(* IEC 61131-3 sources: Industry-PLC-LLM/data/PLCBEAD_repo/PLCBEAD_PLCEmbed-main/PLC-BEAD/Source/OpenPLCv3 (part 4) *)

(* ---- CYCLE_TIME.ST ---- *)
FUNCTION_BLOCK T_PLC_MS_block
	VAR_OUTPUT
		T_PLC_MS :	UDINT;
	END_VAR

	VAR_EXTERNAL
		PLC_TICKS_PER_SEC :	INT;
		PLC_SYS_TICK_CNT :	DINT;
	END_VAR

	VAR
		debug :	BOOL;(*Debug-Mode ON / OFF*)
		N :	INT;(*Debug-Faktor*)
		Offset :	UDINT;(*Debug-Offset*)
		temp :	DWORD := DWORD#1;(*Debug-Offset*)
		mode :	BOOL;(*modus*)
		faktor :	UDINT;(*Systemtakt-Faktor*)
		init :	BOOL;
		v_plc_ticks_per_sec :	UDINT;
		base :	UDINT := UDINT#1000;
	END_VAR

	IF init = FALSE THEN
		v_plc_ticks_per_sec := INT_TO_UDINT(PLC_TICKS_PER_SEC);
		IF v_plc_ticks_per_sec = UDINT#1024 THEN
			faktor := UDINT#1;
			mode := FALSE;
		ELSIF v_plc_ticks_per_sec > UDINT#0 THEN
			IF v_plc_ticks_per_sec <= base THEN
				faktor := base / v_plc_ticks_per_sec;
				mode := FALSE;
			ELSE
				faktor := v_plc_ticks_per_sec / base;
				mode := TRUE;
			END_IF;
		ELSE
			faktor := UDINT#1;
		END_IF;
		init := TRUE;
	END_IF;

	IF mode THEN
		T_PLC_MS := DINT_TO_UDINT(PLC_SYS_TICK_CNT) / faktor;
	ELSE
		T_PLC_MS := DINT_TO_UDINT(PLC_SYS_TICK_CNT) * faktor;
	END_IF;

	IF debug THEN
		T_PLC_MS := (DWORD_TO_UDINT(SHL(UDINT_TO_DWORD(T_PLC_MS),N) OR SHL(temp,N)) - UDINT#1) + Offset;
	END_IF;

END_FUNCTION_BLOCK

FUNCTION_BLOCK CYCLE_TIME
	VAR_INPUT
		RST :	BOOL;
	END_VAR

	VAR_OUTPUT
		CT_MIN :	TIME := t#0s;
		CT_MAX :	TIME := t#0s;
		CT_LAST :	TIME;
		SYSTIME :	TIME;
		SYSDAYS :	INT;
		CYCLES :	DWORD;
	END_VAR

	VAR
		last_cycle :	TIME;
		tx :	TIME;
		init :	BOOL;
		T_PLC_MS :	T_PLC_MS_block;
	END_VAR

	T_PLC_MS();
	tx:= UDINT_TO_TIME(T_PLC_MS.T_PLC_MS) - last_cycle;

	IF rst THEN
		ct_min := t#10h;
		ct_max := t#0ms;
		cycles := DWORD#0;
	ELSIF last_cycle > t#0s THEN
		IF tx < ct_min THEN ct_min := tx;
		ELSIF tx > ct_max THEN ct_max := tx;
		END_IF;
		ct_last := tx;
	ELSIF ct_min = t#0s THEN
		ct_min := t#0s - t#1ms;
	END_IF;
	IF init THEN
		systime := systime + tx;
			IF systime >= t#1d THEN
				systime := systime - t#1d;
				sysdays := sysdays + 1;
			END_IF;
	END_IF;
	init := TRUE;
	last_cycle := last_cycle + tx;
	cycles := UDINT_TO_DWORD(DWORD_TO_UDINT(cycles) + UDINT#1);

END_FUNCTION_BLOCK

PROGRAM program0
  VAR
	RST :	BOOL;

	CT_MIN  :	TIME;
	CT_MAX  :	TIME;
	CT_LAST :	TIME;
	SYSTIME :	TIME;
	SYSDAYS :	INT;
	CYCLES  :	DWORD;

	func_block : CYCLE_TIME;
  END_VAR
	func_block.RST   :=RST ;
	func_block();
	CT_MIN := func_block.CT_MIN ;
	CT_MAX := func_block.CT_MAX ;
	CT_LAST:= func_block.CT_LAST;
	SYSTIME:= func_block.SYSTIME;
	SYSDAYS:= func_block.SYSDAYS;
	CYCLES := func_block.CYCLES ;
END_PROGRAM

CONFIGURATION Config0
	VAR_GLOBAL
		PLC_TICKS_PER_SEC :	INT;
		PLC_SYS_TICK_CNT :	DINT;
	END_VAR

  	RESOURCE Res0 ON PLC
    	TASK task0(INTERVAL := T#20ms,PRIORITY := 0);
    	PROGRAM instance0 WITH task0 : program0;
  	END_RESOURCE
END_CONFIGURATION

(* ---- D_TRIG.ST ---- *)
FUNCTION_BLOCK D_TRIG
	VAR_INPUT
		IN :	DWORD;
	END_VAR

	VAR_OUTPUT
		Q :	BOOL;
		X :	DWORD;
	END_VAR

	VAR
		last_in :	DWORD;
	END_VAR

	Q := in <> last_in;
	X := UDINT_TO_DWORD(DWORD_TO_UDINT(in) - DWORD_TO_UDINT(last_in));
	last_in := in;
END_FUNCTION_BLOCK

PROGRAM program0
  VAR
	IN :	DWORD;

	Q :	BOOL;
	X :	DWORD;

	func_block : D_TRIG;
  END_VAR
	func_block.IN  := IN;
	func_block();
	Q := func_block.Q;
	X := func_block.X;
END_PROGRAM

CONFIGURATION Config0
  RESOURCE Res0 ON PLC
    TASK task0(INTERVAL := T#20ms,PRIORITY := 0);
    PROGRAM instance0 WITH task0 : program0;
  END_RESOURCE
END_CONFIGURATION

(* ---- DATE_TO_STRING.ST ---- *)
FUNCTION YEAR_OF_DATE:INT
	VAR_INPUT
		IDATE :	UDINT;
	END_VAR

	YEAR_OF_DATE := UDINT_TO_INT((idate+UDINT#43200) / UDINT#31557600 + UDINT#1970);
END_FUNCTION

FUNCTION DAY_OF_YEAR:INT
	VAR_INPUT
		IDATE :	UDINT;
	END_VAR

	DAY_OF_YEAR := UDINT_TO_INT(((idate) / UDINT#86400) MOD UDINT#1461);
	IF DAY_OF_YEAR > 729 THEN
		IF DAY_OF_YEAR > 1095 THEN DAY_OF_YEAR := DAY_OF_YEAR - 1095; ELSE DAY_OF_YEAR := DAY_OF_YEAR - 729; END_IF;
	ELSIF DAY_OF_YEAR > 364 THEN
		DAY_OF_YEAR := DAY_OF_YEAR - 364;
	ELSE
		DAY_OF_YEAR := DAY_OF_YEAR + 1;
	END_IF;
END_FUNCTION

FUNCTION LEAP_OF_DATE:BOOL

	VAR_INPUT
		IDATE :	UDINT;
	END_VAR

	LEAP_OF_DATE := SHL(UDINT_TO_DWORD((idate + UDINT#43200) / UDINT#31557600), 30) = DWORD#16#80000000;
END_FUNCTION

FUNCTION MONTH_OF_DATE:INT

	VAR_INPUT
		IDATE :	UDINT;
	END_VAR

	MONTH_OF_DATE := DAY_OF_YEAR(idate);
	IF MONTH_OF_DATE < 32 THEN
		MONTH_OF_DATE := 1;
	ELSIF LEAP_OF_DATE((IDATE)) THEN
		MONTH_OF_DATE := (MONTH_OF_DATE * 53 + 1668) / 1623;
	ELSE
		MONTH_OF_DATE := (MONTH_OF_DATE * 53 + 1700) / 1620;
	END_IF;
END_FUNCTION

FUNCTION DAY_OF_MONTH:INT
	VAR_INPUT
		IDATE :	UDINT;
	END_VAR

	day_of_month := day_of_year(idate);

	IF leap_of_Date((idate)) THEN
		CASE day_of_month OF
			32..60	:	day_of_month := day_of_month - 31;
			61..91	:	day_of_month := day_of_month - 60;
			92..121 :	day_of_month := day_of_month - 91;
			122..152:	day_of_month := day_of_month - 121;
			153..182:	day_of_month := day_of_month - 152;
			183..213:	day_of_month := day_of_month - 182;
			214..244:	day_of_month := day_of_month - 213;
			245..274:	day_of_month := day_of_month - 244;
			275..305:	day_of_month := day_of_month - 274;
			306..335:	day_of_month := day_of_month - 305;
			336..366:	day_of_month := day_of_month - 335;
		END_CASE;
	ELSE
		CASE day_of_month OF
			32..59	:	day_of_month := day_of_month - 31;
			60..90	:	day_of_month := day_of_month - 59;
			91..120 :	day_of_month := day_of_month - 90;
			121..151:	day_of_month := day_of_month - 120;
			152..181:	day_of_month := day_of_month - 151;
			182..212:	day_of_month := day_of_month - 181;
			213..243:	day_of_month := day_of_month - 212;
			244..273:	day_of_month := day_of_month - 243;
			274..304:	day_of_month := day_of_month - 273;
			305..334:	day_of_month := day_of_month - 304;
			335..365:	day_of_month := day_of_month - 334;
		END_CASE;
	END_IF;
END_FUNCTION

FUNCTION_BLOCK DATE_TO_STRING2
	VAR_INPUT
		IDATE :	UDINT;
	END_VAR

	VAR_OUTPUT
		DATE_STRING :	STRING;
	END_VAR

	VAR
		st_tmp1 :	STRING;
	END_VAR

	st_tmp1 := CONCAT(INT_TO_STRING(YEAR_OF_DATE(IDATE)),INT_TO_STRING(MONTH_OF_DATE(IDATE)));
	DATE_STRING := CONCAT(st_tmp1,INT_TO_STRING(day_of_month(IDATE)));
END_FUNCTION_BLOCK

PROGRAM program0
  VAR
    LocalVar0 : UDINT;
	LocalOUT  : STRING;
	func_block : DATE_TO_STRING2;
  END_VAR
	func_block.IDATE  := LocalVar0;
	func_block();
	LocalOUT := func_block.DATE_STRING;
END_PROGRAM

CONFIGURATION Config0
  RESOURCE Res0 ON PLC
    TASK task0(INTERVAL := T#20ms,PRIORITY := 0);
    PROGRAM instance0 WITH task0 : program0;
  END_RESOURCE
END_CONFIGURATION

(* ---- DCF77.ST ---- *)
TYPE
  oscat_dcf77_bits            : ARRAY [0..58]   OF BOOL;
END_TYPE

FUNCTION_BLOCK T_PLC_MS_block
	VAR_OUTPUT
		T_PLC_MS :	UDINT;
	END_VAR

	VAR_EXTERNAL
		PLC_TICKS_PER_SEC :	INT;
		PLC_SYS_TICK_CNT :	DINT;
	END_VAR

	VAR
		debug :	BOOL;(*Debug-Mode ON / OFF*)
		N :	INT;(*Debug-Faktor*)
		Offset :	UDINT;(*Debug-Offset*)
		temp :	DWORD := DWORD#1;(*Debug-Offset*)
		mode :	BOOL;(*modus*)
		faktor :	UDINT;(*Systemtakt-Faktor*)
		init :	BOOL;
		v_plc_ticks_per_sec :	UDINT;
		base :	UDINT := UDINT#1000;
	END_VAR

	IF init = FALSE THEN
		v_plc_ticks_per_sec := INT_TO_UDINT(PLC_TICKS_PER_SEC);
		IF v_plc_ticks_per_sec = UDINT#1024 THEN
			faktor := UDINT#1;
			mode := FALSE;
		ELSIF v_plc_ticks_per_sec > UDINT#0 THEN
			IF v_plc_ticks_per_sec <= base THEN
				faktor := base / v_plc_ticks_per_sec;
				mode := FALSE;
			ELSE
				faktor := v_plc_ticks_per_sec / base;
				mode := TRUE;
			END_IF;
		ELSE
			faktor := UDINT#1;
		END_IF;
		init := TRUE;
	END_IF;

	IF mode THEN
		T_PLC_MS := DINT_TO_UDINT(PLC_SYS_TICK_CNT) / faktor;
	ELSE
		T_PLC_MS := DINT_TO_UDINT(PLC_SYS_TICK_CNT) * faktor;
	END_IF;

	IF debug THEN
		T_PLC_MS := (DWORD_TO_UDINT(SHL(UDINT_TO_DWORD(T_PLC_MS),N) OR SHL(temp,N)) - UDINT#1) + Offset;
	END_IF;

END_FUNCTION_BLOCK

FUNCTION BIT_LOAD_W:WORD
	VAR_INPUT
		IN :	WORD;
		VAL :	BOOL;
		POS :	INT;
	END_VAR

	IF VAL THEN
		BIT_LOAD_W := in OR SHL(WORD#1,pos);
	ELSE
		BIT_LOAD_W := in AND (NOT SHL(WORD#1,pos));
	END_IF;
END_FUNCTION

FUNCTION BIT_OF_DWORD:BOOL
	VAR_INPUT
		IN :	DWORD;
		N :	INT;
	END_VAR
	BIT_OF_DWORD := (SHR(in,n) AND DWORD#1) > DWORD#0;
END_FUNCTION

FUNCTION EVEN:BOOL
	VAR_INPUT
		IN :	DINT;
	END_VAR
	even := NOT BIT_OF_DWORD(DINT_TO_DWORD(in),0);
END_FUNCTION

FUNCTION _INT_TO_UDINT:UDINT
	VAR_INPUT
		IN :	INT;
	END_VAR

	_INT_TO_UDINT := DINT_TO_UDINT(INT_TO_DINT(IN));
END_FUNCTION

FUNCTION SET_DATE:UDINT

	VAR_INPUT
		YEAR :	INT;
		MONTH :	INT;
		DAY :	INT;
	END_VAR

	VAR
		count :	INT;
	END_VAR

	IF month > 2 THEN
		count := (month - 1) * 30;
		IF month > 7 THEN
			count := count + DWORD_TO_INT(SHR(DINT_TO_DWORD(INT_TO_DINT(month) - INT_TO_DINT(3)),1));
		ELSE
			count := count + DWORD_TO_INT(SHR(DINT_TO_DWORD(INT_TO_DINT(month) - INT_TO_DINT(4)),1));
		END_IF;
		IF SHL(INT_TO_WORD(year),14) = WORD#0 THEN
			count := count + 1;
		END_IF;
	ELSE
		count := (month - 1) * 31;
	END_IF;
	SET_DATE := (_INT_TO_UDINT(count + day - 1) + DWORD_TO_UDINT(SHR(UDINT_TO_DWORD(_INT_TO_UDINT(year) * UDINT#1461 - UDINT#2878169), 2))) * UDINT#86400;

END_FUNCTION

FUNCTION DST:BOOL
	VAR_INPUT
		UTC :	UDINT;
	END_VAR

	VAR
		yr :	INT;
		yr4 :	UDINT;
		ltc :	UDINT;
		idate :	UDINT;
	END_VAR

	yr := YEAR_OF_DATE(DT_TO_DATE2(UTC));
	ltc := UTC;
	idate := SET_DT(yr, 3, 31, 1, 0, 0);
	yr4 := DWORD_TO_UDINT(SHR(INT_TO_DWORD(5 * yr), 2)) + UDINT#1;
	DST := (idate - ((yr4 + UDINT#3) MOD UDINT#7) * UDINT#86400 <= ltc) AND (idate + (UDINT#214 - (yr4) MOD UDINT#7) * UDINT#86400 > ltc);

END_FUNCTION

FUNCTION YEAR_OF_DATE:INT
	VAR_INPUT
		IDATE :	UDINT;
	END_VAR

	YEAR_OF_DATE := UDINT_TO_INT((idate+UDINT#43200) / UDINT#31557600 + UDINT#1970);
END_FUNCTION

FUNCTION DAY_OF_WEEK:INT

	VAR_INPUT
		IDATE :	UDINT;
	END_VAR

	DAY_OF_WEEK := UDINT_TO_INT((idate / UDINT#86400 + UDINT#3) MOD UDINT#7) + INT#01;
END_FUNCTION

FUNCTION SET_DT:UDINT
	VAR_INPUT
		YEAR :	INT;
		MONTH :	INT;
		DAY :	INT;
		HOUR :	INT;
		MINUTE :	INT;
		SECOND :	INT;
	END_VAR

	SET_DT := SET_DATE(YEAR, MONTH, DAY) + _INT_TO_UDINT(SECOND) + _INT_TO_UDINT(MINUTE) * UDINT#60 + _INT_TO_UDINT(HOUR) * UDINT#3600;
END_FUNCTION

FUNCTION DT_TO_DATE2:UDINT

	VAR_INPUT
		IN :	UDINT;
	END_VAR

	DT_TO_DATE2 := (IN / UDINT#86400) * UDINT#86400;

END_FUNCTION

FUNCTION_BLOCK DCF77
	VAR_INPUT
		REC :	BOOL;
		SET :	BOOL;
		SDT :	UDINT;
		DSI :	BOOL;
		SYNC_TIMEOUT :	TIME := t#2m;
		TIME_OFFSET :	INT := 1;
		DST_EN :	BOOL := TRUE;
	END_VAR

	VAR_OUTPUT
		TPp :	BOOL;
		DS :	BOOL;
		WDAY :	INT;
		ERROR :	BOOL;
		RTC2 :	UDINT;
		RTC21 :	UDINT;
		MSEC :	INT;
		SYNC :	BOOL;
	END_VAR

	VAR
		MEZ :	UDINT;
		UTC :	UDINT;
		state :	INT;
		edge :	BOOL;
		tx :	TIME;
		ty :	TIME;
		last :	TIME;
		bits :	oscat_dcf77_bits;
		cnt :	INT;
		i :	INT;
		old_time :	UDINT;
		minute :	INT;
		hour :	INT;
		day :	INT;
		month :	INT;
		year :	INT;
		last_sync :	TIME;
		t1 :	TIME;
		tz :	TIME;
		init :	BOOL;
		word_temp :	WORD;
		bool_temp :	BOOL;
		T_PLC_MS :	T_PLC_MS_block;
	END_VAR

	TPp := FALSE;

	T_PLC_MS();
	t1:= UDINT_TO_TIME(T_PLC_MS.T_PLC_MS);
	tx := t1 - last;

	IF rec XOR edge THEN
		edge := rec;
		IF NOT rec AND tx > t#1700ms AND tx < t#2000ms THEN
			(* start condition reached *)
			state := 0;
			tpp := NOT error;
		ELSIF NOT rec AND tx > t#700ms AND tx < t#1000ms THEN
			(* second switch detected *)
			IF state < 58 THEN state := state +1; ELSE state := 0; END_IF;
		ELSIF rec AND tx  < t#120ms THEN
			(* bit 0 detected  *)
			bits[state] := FALSE;
		ELSIF rec AND tx > t#120ms AND tx < t#250ms THEN
			(* bit 1 detected *)
			bits[state] := TRUE;
		ELSE
			(* error condition received signal is not valid *)
			error := TRUE;
			state := 0;
		END_IF;
		last := last + tx;
		IF rec AND state = 58 THEN
			error := FALSE;

			IF bits[0] OR NOT (bits[17] XOR bits[18]) OR NOT bits[20] THEN error := TRUE; END_IF;
			word_temp := WORD#0;

			bool_temp:=bits[21];
			word_temp:=BIT_LOAD_W(word_temp,bool_temp,0);
			bool_temp:=bits[22];
			word_temp:=BIT_LOAD_W(word_temp,bool_temp,1);
			bool_temp:=bits[23];
			word_temp:=BIT_LOAD_W(word_temp,bool_temp,2);
			bool_temp:=bits[24];
			word_temp:=BIT_LOAD_W(word_temp,bool_temp,3);

			minute := WORD_TO_INT(word_temp);
			IF bits[25] THEN minute := minute +10; END_IF;
			IF bits[26] THEN minute := minute +20; END_IF;
			IF bits[27] THEN minute := minute +40; END_IF;
			IF minute > 59 OR (bits[21] XOR bits[22] XOR bits[23] XOR bits[24] XOR bits[25] XOR bits[26] XOR bits[27] XOR bits[28]) THEN error := TRUE; END_IF;

			(* decode hour *)
			word_temp := WORD#0;

			bool_temp:=bits[29];
			word_temp:=BIT_LOAD_W(word_temp,bool_temp,0);    (* word_temp.X0 := bits[29]; *)
			bool_temp:=bits[30];
			word_temp:=BIT_LOAD_W(word_temp,bool_temp,1);    (* word_temp.X1 := bits[30]; *)
			bool_temp:=bits[31];
			word_temp:=BIT_LOAD_W(word_temp,bool_temp,2);    (* word_temp.X2 := bits[31]; *)
			bool_temp:=bits[32];
			word_temp:=BIT_LOAD_W(word_temp,bool_temp,3);    (* word_temp.X3 := bits[32]; *)

			hour := WORD_TO_INT(word_temp);
			IF bits[33] THEN hour := hour +10; END_IF;
			IF bits[34] THEN hour := hour +20; END_IF;
			IF hour > 23 OR (bits[29] XOR bits[30] XOR bits[31] XOR bits[32] XOR bits[33] XOR bits[34] XOR bits[35]) THEN error := TRUE; END_IF;

			(* decode day of month *)
			word_temp := WORD#0;

			bool_temp:=bits[36];
			word_temp:=BIT_LOAD_W(word_temp,bool_temp,0);    (* word_temp.X0 := bits[36]; *)
			bool_temp:=bits[37];
			word_temp:=BIT_LOAD_W(word_temp,bool_temp,1);    (* word_temp.X1 := bits[37]; *)
			bool_temp:=bits[38];
			word_temp:=BIT_LOAD_W(word_temp,bool_temp,2);    (* word_temp.X2 := bits[38]; *)
			bool_temp:=bits[39];
			word_temp:=BIT_LOAD_W(word_temp,bool_temp,3);    (* word_temp.X3 := bits[39]; *)

			day := WORD_TO_INT(word_temp);
			IF bits[40] THEN day := day + 10; END_IF;
			IF bits[41] THEN day := day + 20; END_IF;
			IF day > 31 THEN error := TRUE; END_IF;

			(* decode day of week *)
			word_temp := WORD#0;

			bool_temp:=bits[42];
			word_temp:=BIT_LOAD_W(word_temp,bool_temp,0);    (* word_temp.X0 := bits[42]; *)
			bool_temp:=bits[43];
			word_temp:=BIT_LOAD_W(word_temp,bool_temp,1);    (* word_temp.X1 := bits[43]; *)
			bool_temp:=bits[44];
			word_temp:=BIT_LOAD_W(word_temp,bool_temp,2);    (* word_temp.X2 := bits[44]; *)

			wday := WORD_TO_INT(word_temp);
			IF wday > 7 OR wday < 1 THEN error := TRUE; END_IF;

			(* decode month *)
			word_temp := WORD#0;

			bool_temp:=bits[45];
			word_temp:=BIT_LOAD_W(word_temp,bool_temp,0);    (* word_temp.X0 := bits[45]; *)
			bool_temp:=bits[46];
			word_temp:=BIT_LOAD_W(word_temp,bool_temp,1);    (* word_temp.X1 := bits[46]; *)
			bool_temp:=bits[47];
			word_temp:=BIT_LOAD_W(word_temp,bool_temp,2);    (* word_temp.X2 := bits[47]; *)
			bool_temp:=bits[48];
			word_temp:=BIT_LOAD_W(word_temp,bool_temp,3);    (* word_temp.X3 := bits[48]; *)

			month := WORD_TO_INT(word_temp);
			IF bits[49] THEN month := month +10; END_IF;
			IF month > 12 THEN error := TRUE; END_IF;

			(* decode year *)
			word_temp := WORD#0;

			bool_temp:=bits[50];
			word_temp:=BIT_LOAD_W(word_temp,bool_temp,0);    (* word_temp.X0 := bits[50]; *)
			bool_temp:=bits[51];
			word_temp:=BIT_LOAD_W(word_temp,bool_temp,1);    (* word_temp.X1 := bits[51]; *)
			bool_temp:=bits[52];
			word_temp:=BIT_LOAD_W(word_temp,bool_temp,2);    (* word_temp.X2 := bits[52]; *)
			bool_temp:=bits[53];
			word_temp:=BIT_LOAD_W(word_temp,bool_temp,3);    (* word_temp.X3 := bits[53]; *)

			year := WORD_TO_INT(word_temp);
			IF bits[54] THEN year := year + 10; END_IF;
			IF bits[55] THEN year := year + 20; END_IF;
			IF bits[56] THEN year := year + 40; END_IF;
			IF bits[57] THEN year := year + 80; END_IF;

			(* check parity for bits 36 to 58 *)
			cnt := 0;
			FOR i := 36 TO 58 DO IF bits[i] THEN cnt := cnt + 1; END_IF; END_FOR;
			IF NOT even(INT_TO_DINT(cnt)) THEN error := TRUE; END_IF;

			(* time must be valid for two cycles to clear error flag *)
			IF NOT error THEN
				(* set outputs *)
				old_time := mez;
				IF year >= 70 THEN year := year + 1900; ELSE year := year + 2000; END_IF;
				mez := set_DT(year,month,day,hour,minute,0);
				DS := bits[17];
				IF DS THEN
					UTC := mez - UDINT#7200;
				ELSE
					UTC := mez - UDINT#3600;
				END_IF;

				(* set trigger signal only if the receiver has received 2 successive minutes *)
				IF mez <> old_time + TIME_TO_UDINT(t#1m) THEN error := TRUE ; END_IF;
			END_IF;
		END_IF;
	END_IF;

	tz := UDINT_TO_TIME(_INT_TO_UDINT(ABS(time_offset))* UDINT#3600000);

	IF NOT init OR SET THEN
		init := TRUE;
		utc := sdt;
		tpp := TRUE;
		DS := DSI;
	END_IF;

	IF tpp THEN
		rtc2 := utc;
		IF DS AND dst_en THEN
			IF time_offset < 0 THEN
				rtc21 := rtc2 - TIME_TO_UDINT(tz + t#1h);
			ELSE
				rtc21 := rtc2 + TIME_TO_UDINT(tz + t#1h);
			END_IF;
		ELSE
			IF time_offset < 0 THEN
				rtc21 := rtc2 - TIME_TO_UDINT(tz);
			ELSE
				rtc21 := rtc2 + TIME_TO_UDINT(tz);
			END_IF;
		END_IF;
		sync := TRUE;
		last_sync := last;
		ty := last;
	ELSIF rtc2 > UDINT#0 AND T1 - ty >= t#1s THEN
		rtc2 := rtc2 + TIME_TO_UDINT(t#1s);
		rtc21 := rtc21 + TIME_TO_UDINT(t#1s);
		ty := ty + t#1s;
		sync := ty - last_sync < sync_timeout AND last_sync > t#0s;
		wday := DAY_OF_WEEK(DT_TO_DATE2(rtc21));
		DS := dst_en AND DST(utc);
	END_IF;
	msec := TIME_TO_INT(t1 - ty);

END_FUNCTION_BLOCK

PROGRAM program0
  VAR
	REC         :	BOOL;
	SET         :	BOOL;
	SDT         :	UDINT;
	DSI         :	BOOL;
	SYNC_TIMEOUT:	TIME;
	TIME_OFFSET :	INT;
	DST_EN 	    :	BOOL;

	TPp   :	BOOL;
	DS   :	BOOL;
	WDAY :	INT;
	ERROR:	BOOL;
	RTC2  :	UDINT;
	RTC21 :	UDINT;
	MSEC :	INT;
	SYNC :	BOOL;

	func_block : DCF77;
  END_VAR
	func_block.REC           :=REC         ;
	func_block.SET           :=SET         ;
	func_block.SDT           :=SDT         ;
	func_block.DSI           :=DSI         ;
	func_block.SYNC_TIMEOUT  :=SYNC_TIMEOUT;
	func_block.TIME_OFFSET   :=TIME_OFFSET ;
	func_block.DST_EN 	      :=DST_EN 	    ;
	func_block();
	TPp   := func_block.TPp   ;
	DS   := func_block.DS   ;
	WDAY := func_block.WDAY ;
	ERROR:= func_block.ERROR;
	RTC2  := func_block.RTC2  ;
	RTC21 := func_block.RTC21 ;
	MSEC := func_block.MSEC ;
	SYNC := func_block.SYNC ;
END_PROGRAM

CONFIGURATION Config0
	VAR_GLOBAL
		PLC_TICKS_PER_SEC :	INT;
		PLC_SYS_TICK_CNT :	DINT;
	END_VAR

  	RESOURCE Res0 ON PLC
    	TASK task0(INTERVAL := T#20ms,PRIORITY := 0);
    	PROGRAM instance0 WITH task0 : program0;
  	END_RESOURCE
END_CONFIGURATION

(* ---- DEAD_BAND_A.ST ---- *)
FUNCTION_BLOCK T_PLC_US_Block

	VAR_OUTPUT
		T_PLC_US :	UDINT;
	END_VAR

	VAR_EXTERNAL
		PLC_TICKS_PER_SEC :	INT;
		PLC_SYS_TICK_CNT :	DINT;
	END_VAR

	VAR
		debug :	BOOL;
		N :	INT;
		Offset :	UDINT;
		temp :	DWORD := DWORD#1;
		mode :	BOOL;
		faktor :	UDINT;
		init :	BOOL;
		v_plc_ticks_per_sec :	UDINT;
		base :	UDINT := UDINT#1000000;
	END_VAR

	IF init = FALSE THEN
		v_plc_ticks_per_sec := INT_TO_UDINT(PLC_TICKS_PER_SEC);
		IF v_plc_ticks_per_sec = UDINT#1024 THEN
			faktor := UDINT#1000;
			mode := FALSE;
		ELSIF v_plc_ticks_per_sec > UDINT#0 THEN
			IF v_plc_ticks_per_sec <= base THEN
				faktor := base / v_plc_ticks_per_sec;
				mode := FALSE;
			ELSE
				faktor := v_plc_ticks_per_sec / base;
				mode := TRUE;
			END_IF;
		ELSE
			faktor := UDINT#1;
		END_IF;
		init := TRUE;
	END_IF;

	IF mode THEN
		T_PLC_US := DINT_TO_UDINT(PLC_SYS_TICK_CNT) / faktor;
	ELSE
		T_PLC_US := DINT_TO_UDINT(PLC_SYS_TICK_CNT) * faktor;
	END_IF;

	IF debug THEN
		T_PLC_US := (DWORD_TO_UDINT(SHL(UDINT_TO_DWORD(T_PLC_US),N) OR SHL(temp,N)) - UDINT#1) + Offset;
	END_IF;
END_FUNCTION_BLOCK

FUNCTION_BLOCK FT_PT1

	VAR_INPUT
		IN :	REAL;
		T :	TIME;
		K :	REAL := 1.0;
	END_VAR

	VAR_OUTPUT
		OUT :	REAL;
	END_VAR

	VAR
		last :	UDINT;
		tx :	UDINT;
		init :	BOOL;
		T_PLC_US :	T_PLC_US_Block;
	END_VAR

	T_PLC_US();
	tx:= T_PLC_US.T_PLC_US;

	IF NOT init OR T = t#0s THEN
		init := TRUE;
		out := K * in;
	ELSE
		out := out + (in * K - out) * UDINT_TO_REAL(Tx - last) / TIME_TO_REAL(T) * 1.0E-3;
		IF ABS(out) < 1.0E-20 THEN out := 0.0; END_IF;
	END_IF;
	last := tx;
END_FUNCTION_BLOCK

FUNCTION _REAL_TO_DWORD: DWORD

  VAR_INPUT
    X :	REAL;
  END_VAR

  IF REAL_TO_DWORD(0.5) = DWORD#1 THEN
    _REAL_TO_DWORD := REAL_TO_DWORD(x);
  ELSIF X > 0.0 THEN
    _REAL_TO_DWORD := REAL_TO_DWORD(x+0.5);
  ELSIF X < 0.0 THEN
    _REAL_TO_DWORD := REAL_TO_DWORD(x-0.5);
  ELSE
    _REAL_TO_DWORD := DWORD#0;
  END_IF;
END_FUNCTION

FUNCTION _DWORD_TO_REAL:REAL
	VAR_INPUT
		IN :	DWORD;
	END_VAR

	_DWORD_TO_REAL := UDINT_TO_REAL(DWORD_TO_UDINT(IN));
END_FUNCTION

FUNCTION MULTIME:TIME
	VAR_INPUT
		T :	TIME;
		M :	REAL;
	END_VAR

	multime := DWORD_TO_TIME(_REAL_TO_DWORD(_DWORD_TO_REAL(TIME_TO_DWORD(t))*M));
END_FUNCTION

FUNCTION_BLOCK DEAD_BAND_A
	VAR_INPUT
		X :	REAL;
		T :	TIME;
		KL :	REAL := 1.0;
		LM :	REAL;
	END_VAR

	VAR_OUTPUT
		Y :	REAL;
		L :	REAL;
	END_VAR

	VAR
		tp1 :	FT_PT1;
		tp2 :	FT_PT1;
	END_VAR

	tp1(in := X, T:= T);
	tp2(in := ABS(tp1.out - X), T := MULTIME(T, 4.0));
	L := MIN(KL * tp2.out, LM);

	IF X > L THEN
		Y := X - L;
	ELSIF X < -L THEN
		Y := X + L;
	ELSE
		Y := 0.0;
	END_IF;
END_FUNCTION_BLOCK

PROGRAM program0
  VAR

		X  :	REAL;
		T  :	TIME;
		KL :	REAL;
		LM :	REAL;

		Y :	REAL;
		L :	REAL;

	func_block : DEAD_BAND_A;
  END_VAR
	func_block.X   :=X ;
	func_block.T   :=T ;
	func_block.KL  :=KL;
	func_block.LM  :=LM;
	func_block();
	Y := func_block.Y;
	L := func_block.L;
END_PROGRAM

CONFIGURATION Config0

	VAR_GLOBAL
		PLC_TICKS_PER_SEC :	INT;
		PLC_SYS_TICK_CNT :	DINT;
	END_VAR

	RESOURCE Res0 ON PLC
		TASK task0(INTERVAL := T#20ms,PRIORITY := 0);
		PROGRAM instance0 WITH task0 : program0;
	END_RESOURCE

END_CONFIGURATION

(* ---- DEAD_ZONE2.ST ---- *)
FUNCTION_BLOCK DEAD_ZONE2
	VAR_INPUT
		X :	REAL;
		L :	REAL;
	END_VAR

	VAR_OUTPUT
		Y :	REAL;
	END_VAR

	IF ABS(x) > L THEN
		Y := X;
	ELSIF Y > 0.0 THEN
		Y := L;
	ELSE
		Y := -L;
	END_IF;
END_FUNCTION_BLOCK

PROGRAM program0
  VAR
    LocalVar0 : REAL;
	LocalVar1 : REAL;
	LocalOUT  : REAL;
	func_block : DEAD_ZONE2;
  END_VAR
	func_block.X  := LocalVar0;
	func_block.L  := LocalVar1;
	func_block();
	LocalOUT := func_block.Y;
END_PROGRAM

CONFIGURATION Config0
  RESOURCE Res0 ON PLC
    TASK task0(INTERVAL := T#20ms,PRIORITY := 0);
    PROGRAM instance0 WITH task0 : program0;
  END_RESOURCE
END_CONFIGURATION

(* ---- DEBOUNCE.ST ---- *)
FUNCTION_BLOCK DEBOUNCE_Block

	VAR_INPUT
		IN :	BOOL;
		TD :	TIME;
		PM :	BOOL;
	END_VAR

	VAR_OUTPUT
		Q :	BOOL;
	END_VAR

	VAR
		deb :	TOF;
	END_VAR

	IF NOT deb.Q AND IN THEN
		Q := TRUE;
	ELSIF NOT PM THEN
		Q := deb.Q;
	ELSE
		Q := FALSE;
	END_IF;

END_FUNCTION_BLOCK

PROGRAM program0
	VAR
		IN :	BOOL;
		TD :	TIME;
		PM :	BOOL;
		Q :	BOOL;

		func_block : DEBOUNCE_Block;
	END_VAR
	func_block.IN := IN;
	func_block.TD := TD;
	func_block.PM := PM ;

	func_block();
	Q  := func_block.Q;
END_PROGRAM

CONFIGURATION Config0
	RESOURCE Res0 ON PLC
		TASK task0(INTERVAL := T#20ms,PRIORITY := 0);
		PROGRAM instance0 WITH task0 : program0;
	END_RESOURCE
END_CONFIGURATION

(* ---- DEC_2.ST ---- *)
FUNCTION_BLOCK DEC_2
	VAR_INPUT
		D :	BOOL;
		A :	BOOL;
	END_VAR
	VAR_OUTPUT
		Q0 :	BOOL;
		Q1 :	BOOL;
	END_VAR
	Q0 := D AND NOT A;
	Q1 := D AND A;
END_FUNCTION_BLOCK

PROGRAM program0
  VAR
    LocalVar0 : BOOL;
	LocalVar1 : BOOL;
	LocalOUT  : BOOL;
	LocalOUT1  : BOOL;
	func_block : DEC_2;
  END_VAR
	func_block.D  := LocalVar0;
	func_block.A  := LocalVar1;
	func_block();
	LocalOUT := func_block.Q0;
	LocalOUT1 := func_block.Q1;
END_PROGRAM

CONFIGURATION Config0
  RESOURCE Res0 ON PLC
    TASK task0(INTERVAL := T#20ms,PRIORITY := 0);
    PROGRAM instance0 WITH task0 : program0;
  END_RESOURCE
END_CONFIGURATION

(* ---- DEC_4.ST ---- *)
FUNCTION_BLOCK DEC_4
	VAR_INPUT
		D :	BOOL;
		A0 :	BOOL;
		A1 :	BOOL;
	END_VAR

	VAR_OUTPUT
		Q0 :	BOOL;
		Q1 :	BOOL;
		Q2 :	BOOL;
		Q3 :	BOOL;
	END_VAR

	Q0 := D AND NOT A0 AND NOT A1;
	Q1 := D AND A0 AND NOT A1;
	Q2 := D AND NOT A0 AND A1;
	Q3 := D AND A0 AND A1;
END_FUNCTION_BLOCK

PROGRAM program0
  VAR
	D :	BOOL;
	A0 :	BOOL;
	A1 :	BOOL;

	Q0 :	BOOL;
	Q1 :	BOOL;
	Q2 :	BOOL;
	Q3 :	BOOL;

	func_block : DEC_4;
  END_VAR
	func_block.D   := D  ;
	func_block.A0  := A0  ;
	func_block.A1  := A1  ;
	func_block();
	Q0:= func_block.Q0;
	Q1:= func_block.Q1;
	Q2:= func_block.Q2;
	Q3:= func_block.Q3;
END_PROGRAM

CONFIGURATION Config0
  RESOURCE Res0 ON PLC
    TASK task0(INTERVAL := T#20ms,PRIORITY := 0);
    PROGRAM instance0 WITH task0 : program0;
  END_RESOURCE
END_CONFIGURATION

(* ---- DEC_8.ST ---- *)
FUNCTION BIT_LOAD_B:BYTE
	VAR_INPUT
		IN :	BYTE;
		VAL :	BOOL;
		POS :	INT;
	END_VAR

	IF VAL THEN
		BIT_LOAD_B := in OR SHL(BYTE#1,pos);
	ELSE
		BIT_LOAD_B := in AND (NOT SHL(BYTE#1,pos));
	END_IF;
END_FUNCTION

FUNCTION _BYTE_TO_INT:INT
	VAR_INPUT
		IN :	BYTE;
	END_VAR

	_BYTE_TO_INT := USINT_TO_INT(BYTE_TO_USINT(IN));
END_FUNCTION

FUNCTION_BLOCK DEC_8

	VAR_INPUT
		D :	BOOL;
		A0 :	BOOL;
		A1 :	BOOL;
		A2 :	BOOL;
	END_VAR

	VAR_OUTPUT
		Q0 :	BOOL;
		Q1 :	BOOL;
		Q2 :	BOOL;
		Q3 :	BOOL;
		Q4 :	BOOL;
		Q5 :	BOOL;
		Q6 :	BOOL;
		Q7 :	BOOL;
	END_VAR

	VAR
		X :	BYTE;
	END_VAR

	X:=BIT_LOAD_B(X,A0,0); (* X.0 := A0; *)
	X:=BIT_LOAD_B(X,A1,1); (* X.1 := A1; *)
	X:=BIT_LOAD_B(X,A2,2); (* X.2 := A2; *)

	Q0 := FALSE;
	Q1 := FALSE;
	Q2 := FALSE;
	Q3 := FALSE;
	Q4 := FALSE;
	Q5 := FALSE;
	Q6 := FALSE;
	Q7 := FALSE;

	CASE _BYTE_TO_INT(X) OF
		0 : Q0 := D;
		1 : Q1 := D;
		2 : Q2 := D;
		3 : Q3 := D;
		4 : Q4 := D;
		5 : Q5 := D;
		6 : Q6 := D;
		7 : Q7 := D;
	END_CASE;

	END_FUNCTION_BLOCK

PROGRAM program0
  VAR
	D :	BOOL;
	A0 :	BOOL;
	A1 :	BOOL;
	A2 :	BOOL;

	Q0 :	BOOL;
	Q1 :	BOOL;
	Q2 :	BOOL;
	Q3 :	BOOL;
	Q4 :	BOOL;
	Q5 :	BOOL;
	Q6 :	BOOL;
	Q7 :	BOOL;

	func_block : DEC_8;
  END_VAR
	func_block.D   := D  ;
	func_block.A0  := A0  ;
	func_block.A1  := A1  ;
	func_block.A2  := A2  ;
	func_block();
	Q0:= func_block.Q0;
	Q1:= func_block.Q1;
	Q2:= func_block.Q2;
	Q3:= func_block.Q3;
	Q4:= func_block.Q4;
	Q5:= func_block.Q5;
	Q6:= func_block.Q6;
	Q7:= func_block.Q7;
END_PROGRAM

CONFIGURATION Config0
  RESOURCE Res0 ON PLC
    TASK task0(INTERVAL := T#20ms,PRIORITY := 0);
    PROGRAM instance0 WITH task0 : program0;
  END_RESOURCE
END_CONFIGURATION

(* ---- DEG_TO_DIR.ST ---- *)
TYPE oscat_LANGUAGE:
  STRUCT
    DEFAULT 	: INT;
	LMAX    	: INT;
  END_STRUCT;
END_TYPE

TYPE
  oscat_ELEMENT_DIRS 		: ARRAY [0..15] OF STRING;
  oscat_DIRS				: ARRAY [1..3]  OF oscat_ELEMENT_DIRS := [0,0 , 0];
END_TYPE

FUNCTION_BLOCK SETUP_DIRS
	VAR_IN_OUT
		DIRS :	oscat_DIRS;
	END_VAR

	VAR
		init :	BOOL;
	END_VAR

	IF init THEN RETURN; END_IF;
	init := TRUE;

	(* ---- english --- *)
	DIRS[1][00] := 'N';
	DIRS[1][01] := 'NNE';
	DIRS[1][02] := 'NE';
	DIRS[1][03] := 'ENE';
	DIRS[1][04] := 'E';
	DIRS[1][05] := 'ESE';
	DIRS[1][06] := 'SE';
	DIRS[1][07] := 'SSE';
	DIRS[1][08] := 'S';
	DIRS[1][09] := 'SSW';
	DIRS[1][10] := 'SW';
	DIRS[1][11] := 'WSW';
	DIRS[1][12] := 'W';
	DIRS[1][13] := 'WNW';
	DIRS[1][14] := 'NW';
	DIRS[1][15] := 'NNW';

	(* ---- german --- *)
	DIRS[2][00] := 'N';
	DIRS[2][01] := 'NNO';
	DIRS[2][02] := 'NO';
	DIRS[2][03] := 'ONO';
	DIRS[2][04] := 'O';
	DIRS[2][05] := 'OSO';
	DIRS[2][06] := 'SO';
	DIRS[2][07] := 'SSO';
	DIRS[2][08] := 'S';
	DIRS[2][09] := 'SSW';
	DIRS[2][10] := 'SW';
	DIRS[2][11] := 'WSW';
	DIRS[2][12] := 'W';
	DIRS[2][13] := 'WNW';
	DIRS[2][14] := 'NW';
	DIRS[2][15] := 'NNW';

	(* ---- french --- *)
	DIRS[3][00] := 'N';
	DIRS[3][01] := 'NNO';
	DIRS[3][02] := 'NO';
	DIRS[3][03] := 'ONO';
	DIRS[3][04] := 'O';
	DIRS[3][05] := 'OSO';
	DIRS[3][06] := 'SO';
	DIRS[3][07] := 'SSO';
	DIRS[3][08] := 'S';
	DIRS[3][09] := 'SSW';
	DIRS[3][10] := 'SW';
	DIRS[3][11] := 'WSW';
	DIRS[3][12] := 'W';
	DIRS[3][13] := 'WNW';
	DIRS[3][14] := 'NW';
	DIRS[3][15] := 'NNW';
END_FUNCTION_BLOCK

FUNCTION_BLOCK SETUP_LANGUAGE_Block

	VAR_IN_OUT
		LANGUAGE :	oscat_LANGUAGE;
	END_VAR

	VAR
		init :	BOOL;
	END_VAR

	IF init THEN RETURN; END_IF;
	init := TRUE;

	LANGUAGE.DEFAULT  := 1; (* 1=english, 2=german 3=french *)
	LANGUAGE.LMAX := 3;

END_FUNCTION_BLOCK

FUNCTION_BLOCK DEG_TO_DIR_Block
	VAR_INPUT
		DEG :	INT;
		N :	INT;
		L :	INT;
	END_VAR

	VAR_OUTPUT
		DEG_TO_DIR :	STRING;
	END_VAR

	VAR
		ly :	INT;
		y :	INT;
		SETUP_DIRSS :	SETUP_DIRS;
		DIRS :	oscat_DIRS;
		SETUP_LANGUAGE :	SETUP_LANGUAGE_Block;
		LANGUAGE :	oscat_LANGUAGE;
	END_VAR

	SETUP_DIRSS(DIRS:=DIRS);
	DIRS:=SETUP_DIRSS.DIRS;
	SETUP_LANGUAGE(LANGUAGE:=LANGUAGE);
	LANGUAGE:=SETUP_LANGUAGE.LANGUAGE;

	IF L = 0 THEN ly := LANGUAGE.DEFAULT; ELSE ly := MIN(L, LANGUAGE.LMAX); END_IF;
	y := ((WORD_TO_INT(SHL(INT_TO_WORD(DEG),N-1)) + 45) / 90) MOD WORD_TO_INT(SHL(WORD#2,N))* WORD_TO_INT(SHR(WORD#8,N));
	DEG_TO_DIR := DIRS[ly][y];
END_FUNCTION_BLOCK

PROGRAM program0

	VAR
		DEG :	INT;
		N   :	INT;
		L   :	INT;

		DEG_TO_DIR :	STRING;

		func_block : DEG_TO_DIR_Block;
	END_VAR
		func_block.DEG:=DEG;
		func_block.N  :=N  ;
		func_block.L  :=L  ;

		func_block();
		DEG_TO_DIR := func_block.DEG_TO_DIR;

END_PROGRAM

CONFIGURATION Config0

	RESOURCE Res0 ON PLC
		TASK task0(INTERVAL := T#20ms,PRIORITY := 0);
		PROGRAM instance0 WITH task0 : program0;
	END_RESOURCE

END_CONFIGURATION

(* ---- DEL_CHARS.ST ---- *)
FUNCTION_BLOCK DEL_CHARS_Block
	VAR_INPUT
		IN :	STRING;
		CX :	STRING;
	END_VAR

	VAR_OUTPUT
		DEL_CHARS :	STRING;
	END_VAR

	VAR
		pos :	INT;
		stop :	INT;
		char :	STRING;
	END_VAR

	DEL_CHARS := IN;
	stop := LEN(in);
	pos := 1;
	WHILE pos <= stop DO
		char := MID(DEL_CHARS, 1, pos);
		IF FIND(cx,char) > 0 THEN
			DEL_CHARS := DELETE(DEL_CHARS, 1, pos);
			stop := stop - 1;
		ELSE
			pos := pos + 1;
		END_IF;
	END_WHILE;

END_FUNCTION_BLOCK

PROGRAM program0
  VAR
    LocalVar0 : STRING;
	LocalVar1 : STRING;
	LocalOUT  : STRING;
	func_block : DEL_CHARS_Block;
  END_VAR
	func_block.IN := LocalVar0;
	func_block.CX  := LocalVar1;
	func_block();
	LocalOUT := func_block.DEL_CHARS;
END_PROGRAM

CONFIGURATION Config0
  RESOURCE Res0 ON PLC
    TASK task0(INTERVAL := T#20ms,PRIORITY := 0);
    PROGRAM instance0 WITH task0 : program0;
  END_RESOURCE
END_CONFIGURATION

(* ---- DELAY.ST ---- *)
TYPE
	oscat_delay_buf             : ARRAY [0..31]   OF REAL;
END_TYPE

FUNCTION INC1:INT

	VAR_INPUT
		X :	INT;
		N :	INT;
	END_VAR

	IF X >= N - 1 THEN
		INC1 := 0;
	ELSE
		INC1 := X + 1;
	END_IF;
END_FUNCTION

FUNCTION_BLOCK DELAY

	VAR_INPUT
		IN :	REAL;
		N :	INT;
		RST :	BOOL;
	END_VAR

	VAR_OUTPUT
		OUT :	REAL;
	END_VAR

	VAR
		buf :	oscat_delay_buf;
		i :	INT;
		init :	BOOL;
		stop :	INT;
	END_VAR

	stop := LIMIT(0,N,32) - 1;
	IF rst OR NOT init THEN
		init := TRUE;
		FOR i := 0 TO stop DO buf[i] := in; END_FOR;
		out := in;
		i := 0;
	ELSIF stop < 0 THEN
		out := in;
	ELSE
		out := buf[i];
		buf[i] := in;
		i := INC1(i, N);
	END_IF;

END_FUNCTION_BLOCK

PROGRAM program0
  VAR
	IN :	REAL;
	N :	INT;
	RST :	BOOL;
	OUT :	REAL;
	func_block : DELAY;
  END_VAR
	func_block.IN  :=IN;
	func_block.N  :=N;
	func_block.RST  :=RST;
	func_block();
	OUT := func_block.OUT;

END_PROGRAM

CONFIGURATION Config0
	RESOURCE Res0 ON PLC
		TASK task0(INTERVAL := T#20ms,PRIORITY := 0);
		PROGRAM instance0 WITH task0 : program0;
	END_RESOURCE
END_CONFIGURATION

(* ---- DELAY_4.ST ---- *)
FUNCTION_BLOCK DELAY_4

	VAR_INPUT
		IN :	REAL;
	END_VAR

	VAR_OUTPUT
		OUT1 :	REAL;
		OUT2 :	REAL;
		OUT3 :	REAL;
		OUT4 :	REAL;
	END_VAR

	VAR
		temp :	REAL;
	END_VAR

	out4 := out3;
	out3 := out2;
	out2 := out1;
	out1 := temp;
	temp := in;

END_FUNCTION_BLOCK

PROGRAM program0
  VAR
	IN :	REAL;

	OUT1 :	REAL;
	OUT2 :	REAL;
	OUT3 :	REAL;
	OUT4 :	REAL;
	func_block : DELAY_4;
  END_VAR
	func_block.IN  := IN;
	func_block();
	OUT1:= func_block.OUT1;
	OUT2:= func_block.OUT2;
	OUT3:= func_block.OUT3;
	OUT4:= func_block.OUT4;
END_PROGRAM

CONFIGURATION Config0
  RESOURCE Res0 ON PLC
    TASK task0(INTERVAL := T#20ms,PRIORITY := 0);
    PROGRAM instance0 WITH task0 : program0;
  END_RESOURCE
END_CONFIGURATION

(* ---- DIMM_2.ST ---- *)
FUNCTION UDINT_TO_TIME2:TIME

	VAR_INPUT
		IN :	UDINT;
	END_VAR

	UDINT_TO_TIME2 := DINT_TO_TIME(UDINT_TO_DINT(IN));

END_FUNCTION

FUNCTION_BLOCK T_PLC_MS_block
	VAR_OUTPUT
		T_PLC_MS :	UDINT;
	END_VAR

	VAR_EXTERNAL
		PLC_TICKS_PER_SEC :	INT;
		PLC_SYS_TICK_CNT :	DINT;
	END_VAR

	VAR
		debug :	BOOL;(*Debug-Mode ON / OFF*)
		N :	INT;(*Debug-Faktor*)
		Offset :	UDINT;(*Debug-Offset*)
		temp :	DWORD := DWORD#1;(*Debug-Offset*)
		mode :	BOOL;(*modus*)
		faktor :	UDINT;(*Systemtakt-Faktor*)
		init :	BOOL;
		v_plc_ticks_per_sec :	UDINT;
		base :	UDINT := UDINT#1000;
	END_VAR

	IF init = FALSE THEN
		v_plc_ticks_per_sec := INT_TO_UDINT(PLC_TICKS_PER_SEC);
		IF v_plc_ticks_per_sec = UDINT#1024 THEN
			faktor := UDINT#1;
			mode := FALSE;
		ELSIF v_plc_ticks_per_sec > UDINT#0 THEN
			IF v_plc_ticks_per_sec <= base THEN
				faktor := base / v_plc_ticks_per_sec;
				mode := FALSE;
			ELSE
				faktor := v_plc_ticks_per_sec / base;
				mode := TRUE;
			END_IF;
		ELSE
			faktor := UDINT#1;
		END_IF;
		init := TRUE;
	END_IF;

	IF mode THEN
		T_PLC_MS := DINT_TO_UDINT(PLC_SYS_TICK_CNT) / faktor;
	ELSE
		T_PLC_MS := DINT_TO_UDINT(PLC_SYS_TICK_CNT) * faktor;
	END_IF;

	IF debug THEN
		T_PLC_MS := (DWORD_TO_UDINT(SHL(UDINT_TO_DWORD(T_PLC_MS),N) OR SHL(temp,N)) - UDINT#1) + Offset;
	END_IF;

END_FUNCTION_BLOCK

FUNCTION TIME_TO_UDINT2:UDINT
	VAR_INPUT
		X :	TIME;
	END_VAR

	TIME_TO_UDINT2 := DINT_TO_UDINT(TIME_TO_DINT(X));
END_FUNCTION

FUNCTION FRMP_B:BYTE
	VAR_INPUT
		START :	BYTE;
		DIR :	BOOL;
		TD :	TIME;
		TR :	TIME;
	END_VAR

	IF TD < TR THEN
		FRMP_B := MIN(UDINT_TO_BYTE(DWORD_TO_UDINT(SHL(TIME_TO_DWORD(TD), 8)) / TIME_TO_UDINT2(TR)), SEL(DIR, START, USINT_TO_BYTE(USINT#255 - BYTE_TO_USINT(START))));
		IF DIR THEN
			FRMP_B := USINT_TO_BYTE(BYTE_TO_USINT(START) + BYTE_TO_USINT(FRMP_B));
		ELSE
			FRMP_B := USINT_TO_BYTE(BYTE_TO_USINT(START) - BYTE_TO_USINT(FRMP_B));
		END_IF;
	ELSE
		FRMP_B := SEL(DIR, BYTE#0, BYTE#255);
	END_IF;
END_FUNCTION

FUNCTION_BLOCK _RMP_B
	VAR_INPUT
		DIR :	BOOL;
		E :	BOOL := TRUE;
		TR :	TIME;
	END_VAR

	VAR_IN_OUT
		RMP :	BYTE;
	END_VAR

	VAR
		T_PLC_MS :	T_PLC_MS_Block;
		tx :	TIME;
		tl :	TIME;
		tn :	TIME;
		init :	BOOL;
		last_dir :	BOOL;
		start :	BYTE;
	END_VAR

	T_PLC_MS();
	tx := UDINT_TO_TIME(T_PLC_MS.T_PLC_MS);

	IF E AND init AND (dir = last_dir) AND (RMP <> SEL(DIR, BYTE#0, BYTE#255)) AND TR = tn THEN
		RMP := FRMP_B(start, DIR, tx - tl, TR);
	ELSE
		init := TRUE;
		tl := tx;
		tn := tr;
		start := RMP;
	END_IF;
	last_dir := dir;
END_FUNCTION_BLOCK

FUNCTION_BLOCK CLICK_MODE_Block

	VAR_INPUT
		IN :	BOOL;
		T_LONG :	TIME := T#500ms;
	END_VAR

	VAR_OUTPUT
		SINGLE :	BOOL;
		DOUBLE :	BOOL;
		LONG :	BOOL;
		TP_LONG :	BOOL;
	END_VAR

	VAR
		Timer :	TP;
		cnt :	INT;
		last :	BOOL;
	END_VAR

	timer(in := IN, PT := T_LONG);
	single := FALSE;
	double := FALSE;

	IF timer.Q THEN
		IF NOT in AND last THEN	cnt := cnt + 1; END_IF;
	ELSE
		CASE cnt OF
			1 : single := TRUE;
			2 : double := TRUE;
		END_CASE;
		cnt := 0;
	END_IF;
	last := in;
	TP_LONG := NOT timer.Q AND (NOT LONG) AND IN;
	LONG := NOT timer.Q AND in;

END_FUNCTION_BLOCK

FUNCTION_BLOCK DIMM_2_Block

	VAR_INPUT
		SET :	BOOL;
		VAL :	BYTE := BYTE#255;
		I1 :	BOOL;
		I2 :	BOOL;
		RST :	BOOL;
		T_DEBOUNCE :	TIME := T#10ms;
		T_ON_MAX :	TIME := T#0h;
		T_DIMM_START :	TIME := T#1s;
		T_DIMM :	TIME := T#3s;
		MIN_ON :	BYTE := BYTE#50;
		MAX_ON :	BYTE := BYTE#255;
		RST_OUT :	BOOL;
		SOFT_DIMM :	BOOL := TRUE;
		DBL1_TOG :	BOOL;
		DBL2_TOG :	BOOL;
		DBL1_SET :	BOOL;
		DBL2_SET :	BOOL;
		DBL1_POS :	BYTE;
		DBL2_POS :	BYTE;
	END_VAR

	VAR_OUTPUT
		Q :	BOOL;
		D1 :	BOOL;
		D2 :	BOOL;
	END_VAR

	VAR_IN_OUT
		_OUT :	BYTE;
	END_VAR

	VAR
		t1 :	TOF;
		t2 :	TOF;
		dc1 :	CLICK_MODE_Block;
		dc2 :	CLICK_MODE_Block;
		t3 :	TON;
		dim :	_RMP_B;
	END_VAR

	t1(IN := I1, PT := T_DEBOUNCE);
	t2(IN := I2, PT := T_DEBOUNCE);
	dc1(in := t1.Q, T_LONG := T_DIMM_START);
	dc2(in := t2.Q, T_LONG := T_DIMM_START);

	IF RST THEN
		IF RST_OUT THEN _OUT := BYTE#0; END_IF;
		Q := FALSE;
		D1 := FALSE;
		D2 := FALSE;
	ELSIF set THEN
		_OUT := VAL;
		Q := TRUE;
	ELSIF dc1.SINGLE THEN
		_OUT := LIMIT(MAX(MIN_ON,BYTE#1), _OUT, MAX_ON);
		Q := TRUE;
	ELSIF dc2.SINGLE THEN
		Q := FALSE;
	ELSIF dc1.TP_LONG THEN
		IF NOT Q THEN
			_OUT := SEL(SOFT_DIMM, LIMIT(MAX(MIN_ON,BYTE#1), _OUT, MAX_ON), BYTE#1);
		END_IF;
		Q := TRUE;
		dim.DIR := TRUE;
	ELSIF dc2.TP_LONG THEN
		dim.DIR := FALSE;
	END_IF;

	IF NOT DBL1_TOG THEN D1 := FALSE; END_IF;
	IF dc1.DOUBLE THEN
		IF DBL1_SET THEN
			_OUT := DBL1_POS;
			Q := TRUE;
		ELSE
			D1 := NOT D1;
		END_IF;
	END_IF;
	IF NOT DBL2_TOG THEN D2 := FALSE; END_IF;
	IF dc2.DOUBLE THEN
		IF DBL2_SET THEN
			_OUT := DBL2_POS;
			Q := TRUE;
		ELSE
			D2 := NOT D2;
		END_IF;
	END_IF;

	dim(dir := dc2.LONG, e := dc1.LONG OR dc2.LONG , TR := T_DIMM, rmp := _OUT);
	_OUT := dim.RMP;

	IF _OUT = BYTE#0 THEN Q := FALSE; END_IF;

	IF t_ON_MAX > t#0s THEN
		t3(in := q, pt := T_ON_MAX);
		Q := Q XOR t3.Q;
	END_IF;

END_FUNCTION_BLOCK

PROGRAM program0
	VAR
	    SET :	BOOL;
		VAL :	BYTE := BYTE#255;
		I1 :	BOOL;
		I2 :	BOOL;
		RST :	BOOL;
		T_DEBOUNCE :	TIME := T#10ms;
		T_ON_MAX :	TIME := T#0h;
		T_DIMM_START :	TIME := T#1s;
		T_DIMM :	TIME := T#3s;
		MIN_ON :	BYTE := BYTE#50;
		MAX_ON :	BYTE := BYTE#255;
		RST_OUT :	BOOL;
		SOFT_DIMM :	BOOL := TRUE;
		DBL1_TOG :	BOOL;
		DBL2_TOG :	BOOL;
		DBL1_SET :	BOOL;
		DBL2_SET :	BOOL;
		DBL1_POS :	BYTE;
		DBL2_POS :	BYTE;
		_OUT :	BYTE := BYTE#0;
		Q :	BOOL;
		D1 :	BOOL;
		D2 :	BOOL;

		func_block : DIMM_2_Block;
  	END_VAR
	func_block.SET := SET;
	func_block.VAL := VAL;
	func_block.I1 := I1;
	func_block.I2 := I2;
	func_block.RST := RST;
	func_block.T_DEBOUNCE := T_DEBOUNCE;
	func_block.T_ON_MAX := T_ON_MAX;
	func_block.T_DIMM_START := T_DIMM_START;
	func_block.T_DIMM := T_DIMM;
	func_block.MIN_ON := MIN_ON;
	func_block.MAX_ON := MAX_ON;
	func_block.RST_OUT := RST_OUT;
	func_block.SOFT_DIMM := SOFT_DIMM;
	func_block.DBL1_TOG := DBL1_TOG;
	func_block.DBL2_TOG := DBL2_TOG;
	func_block.DBL1_SET := DBL1_SET;
	func_block.DBL2_SET := DBL2_SET;
	func_block.DBL1_POS := DBL1_POS;
	func_block.DBL2_POS := DBL2_POS;
	func_block._OUT := _OUT;

	func_block();
	_OUT := func_block._OUT;
	Q := func_block.Q;
	D1 := func_block.D1;
	D2 := func_block.D2;
END_PROGRAM

CONFIGURATION Config0
	VAR_GLOBAL
		PLC_TICKS_PER_SEC :	INT;
		PLC_SYS_TICK_CNT :	DINT;
	END_VAR
  	RESOURCE Res0 ON PLC
    	TASK task0(INTERVAL := T#20ms,PRIORITY := 0);
    	PROGRAM instance0 WITH task0 : program0;
  	END_RESOURCE
END_CONFIGURATION

(* ---- DIMM_I.ST ---- *)
FUNCTION_BLOCK SW_RECONFIG_Block

	VAR_INPUT
		IN :	BOOL;
		TD :	TIME;
		TR :	TIME;
	END_VAR

	VAR_OUTPUT
		Q :	BOOL;
	END_VAR

	VAR
		T1 :	TON;
		T2 :	TON;
		INV :	BOOL;
	END_VAR

	t1(in := IN, PT := TD);

	IF tr > t#0s THEN
		Q := t1.Q XOR inv;
		T2(in := Q, pt := TR);
		IF T2.Q THEN INV := NOT INV; END_IF;
	ELSE
		Q := t1.Q;
	END_IF;

END_FUNCTION_BLOCK

FUNCTION_BLOCK CLICK_MODE_Block

	VAR_INPUT
		IN :	BOOL;
		T_LONG :	TIME := T#500ms;
	END_VAR

	VAR_OUTPUT
		SINGLE :	BOOL;
		DOUBLE :	BOOL;
		LONG :	BOOL;
		TP_LONG :	BOOL;
	END_VAR

	VAR
		Timer :	TP;
		cnt :	INT;
		last :	BOOL;
	END_VAR

	timer(in := IN, PT := T_LONG);
	single := FALSE;
	double := FALSE;

	IF timer.Q THEN
		IF NOT in AND last THEN	cnt := cnt + 1; END_IF;
	ELSE
		CASE cnt OF
			1 : single := TRUE;
			2 : double := TRUE;
		END_CASE;
		cnt := 0;
	END_IF;
	last := in;
	TP_LONG := NOT timer.Q AND (NOT LONG) AND IN;
	LONG := NOT timer.Q AND in;

END_FUNCTION_BLOCK

FUNCTION UDINT_TO_TIME2:TIME

	VAR_INPUT
		IN :	UDINT;
	END_VAR

	UDINT_TO_TIME2 := DINT_TO_TIME(UDINT_TO_DINT(IN));

END_FUNCTION

FUNCTION_BLOCK T_PLC_MS_block
	VAR_OUTPUT
		T_PLC_MS :	UDINT;
	END_VAR

	VAR_EXTERNAL
		PLC_TICKS_PER_SEC :	INT;
		PLC_SYS_TICK_CNT :	DINT;
	END_VAR

	VAR
		debug :	BOOL;(*Debug-Mode ON / OFF*)
		N :	INT;(*Debug-Faktor*)
		Offset :	UDINT;(*Debug-Offset*)
		temp :	DWORD := DWORD#1;(*Debug-Offset*)
		mode :	BOOL;(*modus*)
		faktor :	UDINT;(*Systemtakt-Faktor*)
		init :	BOOL;
		v_plc_ticks_per_sec :	UDINT;
		base :	UDINT := UDINT#1000;
	END_VAR

	IF init = FALSE THEN
		v_plc_ticks_per_sec := INT_TO_UDINT(PLC_TICKS_PER_SEC);
		IF v_plc_ticks_per_sec = UDINT#1024 THEN
			faktor := UDINT#1;
			mode := FALSE;
		ELSIF v_plc_ticks_per_sec > UDINT#0 THEN
			IF v_plc_ticks_per_sec <= base THEN
				faktor := base / v_plc_ticks_per_sec;
				mode := FALSE;
			ELSE
				faktor := v_plc_ticks_per_sec / base;
				mode := TRUE;
			END_IF;
		ELSE
			faktor := UDINT#1;
		END_IF;
		init := TRUE;
	END_IF;

	IF mode THEN
		T_PLC_MS := DINT_TO_UDINT(PLC_SYS_TICK_CNT) / faktor;
	ELSE
		T_PLC_MS := DINT_TO_UDINT(PLC_SYS_TICK_CNT) * faktor;
	END_IF;

	IF debug THEN
		T_PLC_MS := (DWORD_TO_UDINT(SHL(UDINT_TO_DWORD(T_PLC_MS),N) OR SHL(temp,N)) - UDINT#1) + Offset;
	END_IF;

END_FUNCTION_BLOCK

FUNCTION TIME_TO_UDINT2:UDINT
	VAR_INPUT
		X :	TIME;
	END_VAR

	TIME_TO_UDINT2 := DINT_TO_UDINT(TIME_TO_DINT(X));
END_FUNCTION

FUNCTION FRMP_B:BYTE
	VAR_INPUT
		START :	BYTE;
		DIR :	BOOL;
		TD :	TIME;
		TR :	TIME;
	END_VAR

	IF TD < TR THEN
		FRMP_B := MIN(UDINT_TO_BYTE(DWORD_TO_UDINT(SHL(TIME_TO_DWORD(TD), 8)) / TIME_TO_UDINT2(TR)), SEL(DIR, START, USINT_TO_BYTE(USINT#255 - BYTE_TO_USINT(START))));
		IF DIR THEN
			FRMP_B := USINT_TO_BYTE(BYTE_TO_USINT(START) + BYTE_TO_USINT(FRMP_B));
		ELSE
			FRMP_B := USINT_TO_BYTE(BYTE_TO_USINT(START) - BYTE_TO_USINT(FRMP_B));
		END_IF;
	ELSE
		FRMP_B := SEL(DIR, BYTE#0, BYTE#255);
	END_IF;
END_FUNCTION

FUNCTION_BLOCK _RMP_B
	VAR_INPUT
		DIR :	BOOL;
		E :	BOOL := TRUE;
		TR :	TIME;
	END_VAR

	VAR_IN_OUT
		RMP :	BYTE;
	END_VAR

	VAR
		T_PLC_MS :	T_PLC_MS_block;
		tx :	TIME;
		tl :	TIME;
		tn :	TIME;
		init :	BOOL;
		last_dir :	BOOL;
		start :	BYTE;
	END_VAR

	T_PLC_MS();
	tx := UDINT_TO_TIME(T_PLC_MS.T_PLC_MS);

	IF E AND init AND (dir = last_dir) AND (RMP <> SEL(DIR, BYTE#0, BYTE#255)) AND TR = tn THEN
		RMP := FRMP_B(start, DIR, tx - tl, TR);
	ELSE
		init := TRUE;
		tl := tx;
		tn := tr;
		start := RMP;
	END_IF;
	last_dir := dir;
END_FUNCTION_BLOCK

FUNCTION _BYTE_TO_INT:INT
	VAR_INPUT
		IN :	BYTE;
	END_VAR

	_BYTE_TO_INT := USINT_TO_INT(BYTE_TO_USINT(IN));
END_FUNCTION

FUNCTION_BLOCK DIMM_I_Block

	VAR_INPUT
		SET :	BOOL;
		VAL :	BYTE := BYTE#255;
		IN :	BOOL;
		RST :	BOOL;
		T_DEBOUNCE :	TIME := T#10ms;
		T_RECONFIG :	TIME := T#10s;
		T_ON_MAX :	TIME := T#0h;
		T_DIMM_START :	TIME := T#1s;
		T_DIMM :	TIME := T#3s;
		MIN_ON :	BYTE := BYTE#50;
		MAX_ON :	BYTE := BYTE#255;
		SOFT_DIMM :	BOOL := TRUE;
		DBL_TOGGLE :	BOOL;
		RST_OUT :	BOOL;
	END_VAR

	VAR_OUTPUT
		Q :	BOOL;
		DBL :	BOOL;
	END_VAR

	VAR_IN_OUT
		OUT :	BYTE;
	END_VAR

	VAR
		config :	SW_RECONFIG_Block;
		decode :	CLICK_MODE_Block;
		t3 :	TON;
		dim :	_RMP_B;
		dir :	BOOL;
	END_VAR

	config(IN := IN, TD := T_DEBOUNCE, TR := T_RECONFIG);
	decode(in := config.Q, T_LONG := T_DIMM_START);

	IF RST THEN
		IF rst_out THEN out := BYTE#0; END_IF;
		Q := FALSE;
		dir := out > BYTE#127;
	ELSIF set THEN
		out := val;
		Q := TRUE;
		dir := out > BYTE#127;
	ELSIF decode.SINGLE THEN
		Q := NOT Q;
		IF Q THEN OUT := INT_TO_BYTE(LIMIT_INT(MAX(_BYTE_TO_INT(MIN_ON),1), _BYTE_TO_INT(out), _BYTE_TO_INT(MAX_ON)));	END_IF;
		dir := OUT > BYTE#127;
	ELSIF decode.TP_LONG THEN
		IF NOT Q THEN
			IF SOFT_DIMM THEN
				OUT := BYTE#1;
				dir := TRUE;
			ELSE
				out := INT_TO_BYTE(LIMIT_INT(MAX(_BYTE_TO_INT(MIN_ON),1), _BYTE_TO_INT(out), _BYTE_TO_INT(MAX_ON)));
				DIR := out < BYTE#127;
			END_IF;
			Q := TRUE;
		ELSE
			dir := NOT dir;
		END_IF;
	END_IF;

	IF NOT dbl_toggle THEN dbl := FALSE; END_IF;
	IF decode.DOUBLE THEN dbl := NOT dbl; END_IF;

	dim(DIR := dir, e := decode.LONG AND Q, TR := T_DIMM, rmp := out);
	OUT := dim.RMP;
	IF out = BYTE#0 THEN
		dir := TRUE;
	ELSIF out = BYTE#255 THEN
		dir := FALSE;
	END_IF;

	IF t_ON_MAX > t#0s THEN
		t3(in := q, pt := T_ON_MAX);
		Q := Q XOR t3.Q;
	END_IF;

END_FUNCTION_BLOCK

PROGRAM program0
	VAR
	    SET :	BOOL;
		VAL :	BYTE := BYTE#255;
		IN :	BOOL;
		RST :	BOOL;
		T_DEBOUNCE :	TIME := T#10ms;
		T_RECONFIG :	TIME := T#10s;
		T_ON_MAX :	TIME := T#0h;
		T_DIMM_START :	TIME := T#1s;
		T_DIMM :	TIME := T#3s;
		MIN_ON :	BYTE := BYTE#50;
		MAX_ON :	BYTE := BYTE#255;
		SOFT_DIMM :	BOOL := TRUE;
		DBL_TOGGLE :	BOOL;
		RST_OUT :	BOOL;
		OUT :	BYTE;
		Q :	BOOL;
		DBL :	BOOL;

		func_block : DIMM_I_Block;
  	END_VAR
	func_block.SET := SET;
	func_block.VAL := VAL;
	func_block.IN := IN;
	func_block.RST := RST;
	func_block.T_DEBOUNCE := T_DEBOUNCE;
	func_block.T_RECONFIG := T_RECONFIG;
	func_block.T_ON_MAX := T_ON_MAX;
	func_block.T_DIMM_START := T_DIMM_START;
	func_block.T_DIMM := T_DIMM;
	func_block.MIN_ON := MIN_ON;
	func_block.MAX_ON := MAX_ON;
	func_block.SOFT_DIMM := SOFT_DIMM;
	func_block.DBL_TOGGLE := DBL_TOGGLE;
	func_block.RST_OUT := RST_OUT;
	func_block.OUT := OUT;

	func_block();
	OUT := func_block.OUT;
	Q := func_block.Q;
	DBL := func_block.DBL;
END_PROGRAM

CONFIGURATION Config0
	VAR_GLOBAL
		PLC_TICKS_PER_SEC :	INT;
		PLC_SYS_TICK_CNT :	DINT;
	END_VAR
  	RESOURCE Res0 ON PLC
    	TASK task0(INTERVAL := T#20ms,PRIORITY := 0);
    	PROGRAM instance0 WITH task0 : program0;
  	END_RESOURCE
END_CONFIGURATION

(* ---- DIR_TO_DEG.ST ---- *)
TYPE oscat_LANGUAGE:
  STRUCT
    DEFAULT 	: INT;
	LMAX    	: INT;
  END_STRUCT;
END_TYPE

TYPE
  oscat_ELEMENT_DIRS 		: ARRAY [0..15] OF STRING;
  oscat_DIRS				: ARRAY [1..3]  OF oscat_ELEMENT_DIRS := [0,0 , 0];
END_TYPE

FUNCTION_BLOCK SETUP_DIRS
	VAR_IN_OUT
		DIRS :	oscat_DIRS;
	END_VAR

	VAR
		init :	BOOL;
	END_VAR

	IF init THEN RETURN; END_IF;
	init := TRUE;

	(* ---- english --- *)
	DIRS[1][00] := 'N';
	DIRS[1][01] := 'NNE';
	DIRS[1][02] := 'NE';
	DIRS[1][03] := 'ENE';
	DIRS[1][04] := 'E';
	DIRS[1][05] := 'ESE';
	DIRS[1][06] := 'SE';
	DIRS[1][07] := 'SSE';
	DIRS[1][08] := 'S';
	DIRS[1][09] := 'SSW';
	DIRS[1][10] := 'SW';
	DIRS[1][11] := 'WSW';
	DIRS[1][12] := 'W';
	DIRS[1][13] := 'WNW';
	DIRS[1][14] := 'NW';
	DIRS[1][15] := 'NNW';

	(* ---- german --- *)
	DIRS[2][00] := 'N';
	DIRS[2][01] := 'NNO';
	DIRS[2][02] := 'NO';
	DIRS[2][03] := 'ONO';
	DIRS[2][04] := 'O';
	DIRS[2][05] := 'OSO';
	DIRS[2][06] := 'SO';
	DIRS[2][07] := 'SSO';
	DIRS[2][08] := 'S';
	DIRS[2][09] := 'SSW';
	DIRS[2][10] := 'SW';
	DIRS[2][11] := 'WSW';
	DIRS[2][12] := 'W';
	DIRS[2][13] := 'WNW';
	DIRS[2][14] := 'NW';
	DIRS[2][15] := 'NNW';

	(* ---- french --- *)
	DIRS[3][00] := 'N';
	DIRS[3][01] := 'NNO';
	DIRS[3][02] := 'NO';
	DIRS[3][03] := 'ONO';
	DIRS[3][04] := 'O';
	DIRS[3][05] := 'OSO';
	DIRS[3][06] := 'SO';
	DIRS[3][07] := 'SSO';
	DIRS[3][08] := 'S';
	DIRS[3][09] := 'SSW';
	DIRS[3][10] := 'SW';
	DIRS[3][11] := 'WSW';
	DIRS[3][12] := 'W';
	DIRS[3][13] := 'WNW';
	DIRS[3][14] := 'NW';
	DIRS[3][15] := 'NNW';
END_FUNCTION_BLOCK

FUNCTION_BLOCK SETUP_LANGUAGE_Block

	VAR_IN_OUT
		LANGUAGE :	oscat_LANGUAGE;
	END_VAR

	VAR
		init :	BOOL;
	END_VAR

	IF init THEN RETURN; END_IF;
	init := TRUE;

	LANGUAGE.DEFAULT  := 1; (* 1=english, 2=german 3=french *)
	LANGUAGE.LMAX := 3;

END_FUNCTION_BLOCK

FUNCTION_BLOCK DIR_TO_DEG_Block
	VAR_INPUT
		DIR :	STRING;
		L :	INT;
	END_VAR

	VAR_OUTPUT
		DIR_TO_DEG :	INT;
	END_VAR

	VAR
		ly :	INT;
		i :	INT;
		SETUP_DIRSS :	SETUP_DIRS;
		DIRS :	oscat_DIRS;
		SETUP_LANGUAGE :	SETUP_LANGUAGE_Block;
		LANGUAGE :	oscat_LANGUAGE;
	END_VAR

	SETUP_DIRSS(DIRS:=DIRS);
	DIRS:=SETUP_DIRSS.DIRS;
	SETUP_LANGUAGE(LANGUAGE:=LANGUAGE);
	LANGUAGE:=SETUP_LANGUAGE.LANGUAGE;

	IF L = 0 THEN ly := LANGUAGE.DEFAULT; ELSE ly := MIN(L, LANGUAGE.LMAX); END_IF;
	FOR i := 0 TO 15 DO
		IF EQ_STRING(DIRS[ly][i],DIR) THEN EXIT; END_IF;
	END_FOR;
	DIR_TO_DEG := WORD_TO_INT(SHR(INT_TO_WORD(i * 45 + 1), 1));

END_FUNCTION_BLOCK

PROGRAM program0
  VAR
    LocalVar0 : STRING;
	LocalVar1 : INT;

	LocalOUT  : INT;
	func_block : DIR_TO_DEG_Block;
  END_VAR
	func_block.DIR  := LocalVar0;
	func_block.L  := LocalVar1;
	func_block();
	LocalOUT := func_block.DIR_TO_DEG;
END_PROGRAM

CONFIGURATION Config0
  RESOURCE Res0 ON PLC
    TASK task0(INTERVAL := T#20ms,PRIORITY := 0);
    PROGRAM instance0 WITH task0 : program0;
  END_RESOURCE
END_CONFIGURATION

(* ---- DRIVER_1.ST ---- *)
FUNCTION_BLOCK DRIVER_1
	VAR_INPUT
		SET :	BOOL;
		IN :	BOOL;
		RST :	BOOL;
		TOGGLE_MODE :	BOOL;
		TIMEOUT :	TIME;
	END_VAR

	VAR_OUTPUT
		Q :	BOOL;
	END_VAR

	VAR
		off :	TON;
		edge :	BOOL;
	END_VAR

	IF off.Q THEN Q := FALSE; END_IF;
	IF rst THEN
		Q := FALSE;
	ELSIF set THEN
		Q := TRUE;
	ELSIF IN AND NOT edge THEN
		IF toggle_mode THEN q := NOT Q; ELSE q := TRUE; END_IF;
	END_IF;
	edge := in;
	IF timeout > t#0s THEN off(in := Q, PT := Timeout); END_IF;

END_FUNCTION_BLOCK

PROGRAM program0
  VAR
	SET         :	BOOL;
	IN          :	BOOL;
	RST         :	BOOL;
	TOGGLE_MODE :	BOOL;
	TIMEOUT     :	TIME;

	Q :	BOOL;

	func_block : DRIVER_1;
  END_VAR
	func_block.SET         :=SET        ;
	func_block.IN          :=IN         ;
	func_block.RST         :=RST        ;
	func_block.TOGGLE_MODE :=TOGGLE_MODE;
	func_block.TIMEOUT     :=TIMEOUT    ;
	func_block();
	Q := func_block.Q;
END_PROGRAM

CONFIGURATION Config0
  RESOURCE Res0 ON PLC
    TASK task0(INTERVAL := T#20ms,PRIORITY := 0);
    PROGRAM instance0 WITH task0 : program0;
  END_RESOURCE
END_CONFIGURATION

(* ---- DRIVER_4.ST ---- *)
FUNCTION_BLOCK DRIVER_1
	VAR_INPUT
		SET :	BOOL;
		IN :	BOOL;
		RST :	BOOL;
		TOGGLE_MODE :	BOOL;
		TIMEOUT :	TIME;
	END_VAR

	VAR_OUTPUT
		Q :	BOOL;
	END_VAR

	VAR
		off :	TON;
		edge :	BOOL;
	END_VAR

	IF off.Q THEN Q := FALSE; END_IF;
	IF rst THEN
		Q := FALSE;
	ELSIF set THEN
		Q := TRUE;
	ELSIF IN AND NOT edge THEN
		IF toggle_mode THEN q := NOT Q; ELSE q := TRUE; END_IF;
	END_IF;
	edge := in;
	IF timeout > t#0s THEN off(in := Q, PT := Timeout); END_IF;

END_FUNCTION_BLOCK

FUNCTION_BLOCK DRIVER_4

	VAR_INPUT
		SET :	BOOL;
		IN0 :	BOOL;
		IN1 :	BOOL;
		IN2 :	BOOL;
		IN3 :	BOOL;
		RST :	BOOL;
		TOGGLE_MODE :	BOOL;
		TIMEOUT :	TIME;
	END_VAR

	VAR_OUTPUT
		Q0 :	BOOL;
		Q1 :	BOOL;
		Q2 :	BOOL;
		Q3 :	BOOL;
	END_VAR

	VAR
		d0 :	DRIVER_1;
		d1 :	DRIVER_1;
		d2 :	DRIVER_1;
		d3 :	DRIVER_1;
	END_VAR

	D0(Set:=set, in:=in0, rst:=rst, toggle_mode:=toggle_mode, timeout:=timeout);
	D1(Set:=set, in:=in1, rst:=rst, toggle_mode:=toggle_mode, timeout:=timeout);
	D2(Set:=set, in:=in2, rst:=rst, toggle_mode:=toggle_mode, timeout:=timeout);
	D3(Set:=set, in:=in3, rst:=rst, toggle_mode:=toggle_mode, timeout:=timeout);
	Q0 := D0.Q;
	Q1 := D1.Q;
	Q2 := D2.Q;
	Q3 := D3.Q;

END_FUNCTION_BLOCK

PROGRAM program0
  VAR
	SET         :	BOOL;
	IN0         :	BOOL;
	IN1         :	BOOL;
	IN2         :	BOOL;
	IN3         :	BOOL;
	RST         :	BOOL;
	TOGGLE_MODE :	BOOL;
	TIMEOUT     :	TIME;

	Q0 :	BOOL;
	Q1 :	BOOL;
	Q2 :	BOOL;
	Q3 :	BOOL;

	func_block : DRIVER_4;
  END_VAR
	func_block.SET         := SET        ;
	func_block.IN0         := IN0        ;
	func_block.IN1         := IN1        ;
	func_block.IN2         := IN2        ;
	func_block.IN3         := IN3        ;
	func_block.RST         := RST        ;
	func_block.TOGGLE_MODE := TOGGLE_MODE;
	func_block.TIMEOUT     := TIMEOUT    ;
	func_block();
	Q0 := func_block.Q0;
	Q1 := func_block.Q1;
	Q2 := func_block.Q2;
	Q3 := func_block.Q3;
END_PROGRAM

CONFIGURATION Config0
  RESOURCE Res0 ON PLC
    TASK task0(INTERVAL := T#20ms,PRIORITY := 0);
    PROGRAM instance0 WITH task0 : program0;
  END_RESOURCE
END_CONFIGURATION

(* ---- DRIVER_4C.ST ---- *)
TYPE
  oscat_DRIVER_4C 			  : ARRAY [1..7] 	OF BYTE;
END_TYPE
FUNCTION_BLOCK DRIVER_4C

	VAR_INPUT
		IN :	BOOL;
		RST :	BOOL;
		TIMEOUT :	TIME;
		SX :	oscat_DRIVER_4C;
	END_VAR

	VAR_OUTPUT
		SN :	INT;
		Q0 :	BOOL;
		Q1 :	BOOL;
		Q2 :	BOOL;
		Q3 :	BOOL;
	END_VAR

	VAR
		off :	TON;
		edge :	BOOL;
	END_VAR

	IF RST OR off.Q THEN
		SN := 0;
	ELSIF IN AND NOT edge THEN
		SN := SN + 1;
		IF SN > 7 OR SX[SN] = BYTE#0 THEN SN := 0; END_IF;
	END_IF;
	edge := in;
	IF SN > 0 THEN
		Q0 := (SX[SN] AND BYTE#1) > BYTE#0;
		Q1 := (SX[SN] AND BYTE#2) > BYTE#0;
		Q2 := (SX[SN] AND BYTE#4) > BYTE#0;
		Q3 := (SX[SN] AND BYTE#8) > BYTE#0;
	ELSE
		Q0 := FALSE;
		Q1 := FALSE;
		Q2 := FALSE;
		Q3 := FALSE;
	END_IF;

	IF timeout > t#0s THEN off(in := SN > 0, PT := Timeout); END_IF;

END_FUNCTION_BLOCK

PROGRAM program0
  VAR
	IN      :	BOOL;
	RST     :	BOOL;
	TIMEOUT :	TIME;
	SX      :	oscat_DRIVER_4C;

	SN :	INT;
	Q0 :	BOOL;
	Q1 :	BOOL;
	Q2 :	BOOL;
	Q3 :	BOOL;

	func_block : DRIVER_4C;
  END_VAR
	func_block.IN       :=IN      ;
	func_block.RST      :=RST     ;
	func_block.TIMEOUT  :=TIMEOUT ;
	func_block.SX       :=SX      ;
	func_block();
	SN := func_block.SN;
	Q0 := func_block.Q0;
	Q1 := func_block.Q1;
	Q2 := func_block.Q2;
	Q3 := func_block.Q3;
END_PROGRAM

CONFIGURATION Config0
  RESOURCE Res0 ON PLC
    TASK task0(INTERVAL := T#20ms,PRIORITY := 0);
    PROGRAM instance0 WITH task0 : program0;
  END_RESOURCE
END_CONFIGURATION

(* ---- DT2_TO_SDT.ST ---- *)
TYPE oscat_SDT :
STRUCT
	YEAR : INT;
	MONTH : INT;
	DAY : INT;
	WEEKDAY : INT;
	HOUR : INT;
	MINUTE : INT;
	SECOND : INT;
	MS : INT;
END_STRUCT;
END_TYPE

FUNCTION DAY_OF_WEEK:INT

	VAR_INPUT
		IDATE :	UDINT;
	END_VAR

	DAY_OF_WEEK := UDINT_TO_INT((idate / UDINT#86400 + UDINT#3) MOD UDINT#7) + INT#01;
END_FUNCTION

FUNCTION DAY_OF_YEAR:INT
	VAR_INPUT
		IDATE :	UDINT;
	END_VAR

	DAY_OF_YEAR := UDINT_TO_INT(((idate) / UDINT#86400) MOD UDINT#1461);
	IF DAY_OF_YEAR > 729 THEN
		IF DAY_OF_YEAR > 1095 THEN DAY_OF_YEAR := DAY_OF_YEAR - 1095; ELSE DAY_OF_YEAR := DAY_OF_YEAR - 729; END_IF;
	ELSIF DAY_OF_YEAR > 364 THEN
		DAY_OF_YEAR := DAY_OF_YEAR - 364;
	ELSE
		DAY_OF_YEAR := DAY_OF_YEAR + 1;
	END_IF;
END_FUNCTION

FUNCTION LEAP_OF_DATE:BOOL

	VAR_INPUT
		IDATE :	UDINT;
	END_VAR

	LEAP_OF_DATE := SHL(UDINT_TO_DWORD((idate + UDINT#43200) / UDINT#31557600), 30) = DWORD#16#80000000;
END_FUNCTION

FUNCTION DAY_OF_MONTH:INT
	VAR_INPUT
		IDATE :	UDINT;
	END_VAR

	day_of_month := day_of_year(idate);

	IF leap_of_Date(idate) THEN
		CASE day_of_month OF
			32..60	:	day_of_month := day_of_month - 31;
			61..91	:	day_of_month := day_of_month - 60;
			92..121 :	day_of_month := day_of_month - 91;
			122..152:	day_of_month := day_of_month - 121;
			153..182:	day_of_month := day_of_month - 152;
			183..213:	day_of_month := day_of_month - 182;
			214..244:	day_of_month := day_of_month - 213;
			245..274:	day_of_month := day_of_month - 244;
			275..305:	day_of_month := day_of_month - 274;
			306..335:	day_of_month := day_of_month - 305;
			336..366:	day_of_month := day_of_month - 335;
		END_CASE;
	ELSE
		CASE day_of_month OF
			32..59	:	day_of_month := day_of_month - 31;
			60..90	:	day_of_month := day_of_month - 59;
			91..120 :	day_of_month := day_of_month - 90;
			121..151:	day_of_month := day_of_month - 120;
			152..181:	day_of_month := day_of_month - 151;
			182..212:	day_of_month := day_of_month - 181;
			213..243:	day_of_month := day_of_month - 212;
			244..273:	day_of_month := day_of_month - 243;
			274..304:	day_of_month := day_of_month - 273;
			305..334:	day_of_month := day_of_month - 304;
			335..365:	day_of_month := day_of_month - 334;
		END_CASE;
	END_IF;
END_FUNCTION

FUNCTION MONTH_OF_DATE:INT

	VAR_INPUT
		IDATE :	UDINT;
	END_VAR

	MONTH_OF_DATE := DAY_OF_YEAR(idate);
	IF MONTH_OF_DATE < 32 THEN
		MONTH_OF_DATE := 1;
	ELSIF LEAP_OF_DATE((IDATE)) THEN
		MONTH_OF_DATE := (MONTH_OF_DATE * 53 + 1668) / 1623;
	ELSE
		MONTH_OF_DATE := (MONTH_OF_DATE * 53 + 1700) / 1620;
	END_IF;
END_FUNCTION

FUNCTION YEAR_OF_DATE:INT
	VAR_INPUT
		IDATE :	UDINT;
	END_VAR

	YEAR_OF_DATE := UDINT_TO_INT((idate+UDINT#43200) / UDINT#31557600 + UDINT#1970);
END_FUNCTION

FUNCTION_BLOCK DT2_TO_SDT
VAR_INPUT
	DI :	UDINT;
	TI :	UDINT;
END_VAR

VAR_OUTPUT
	SDT :	oscat_SDT;
END_VAR

SDT.YEAR := YEAR_OF_DATE(di);
SDT.MONTH := MONTH_OF_DATE(di);
SDT.DAY := DAY_OF_MONTH(di);
SDT.WEEKDAY := DAY_OF_WEEK(di);
SDT.MS := UDINT_TO_INT(ti MOD UDINT#1000);
SDT.SECOND := UDINT_TO_INT((ti / UDINT#1000) MOD UDINT#60);
SDT.MINUTE := UDINT_TO_INT((ti / UDINT#60000) MOD UDINT#60);
SDT.HOUR := UDINT_TO_INT(ti / UDINT#3600000);

END_FUNCTION_BLOCK

PROGRAM program0
  VAR
    LocalVar0 : UDINT;
	LocalVar1 : UDINT;
	LocalOUT  : oscat_SDT;
	func_block : DT2_TO_SDT;
  END_VAR
	func_block.DI  := LocalVar0;
	func_block.TI  := LocalVar1;
	func_block();
	LocalOUT := func_block.SDT;
END_PROGRAM

CONFIGURATION Config0
  RESOURCE Res0 ON PLC
    TASK task0(INTERVAL := T#20ms,PRIORITY := 0);
    PROGRAM instance0 WITH task0 : program0;
  END_RESOURCE
END_CONFIGURATION

(* ---- DT_SIMU.ST ---- *)
FUNCTION _REAL_TO_UDINT:UDINT
  VAR_INPUT
    X :	REAL;
  END_VAR

  IF REAL_TO_UDINT(0.5) = UDINT#1 THEN
    _REAL_TO_UDINT := REAL_TO_UDINT(x);
  ELSIF X > 0.0 THEN
    _REAL_TO_UDINT := REAL_TO_UDINT(x+0.5);
  ELSIF X < 0.0 THEN
    _REAL_TO_UDINT := REAL_TO_UDINT(x-0.5);
  ELSE
    _REAL_TO_UDINT := UDINT#0;
  END_IF;
END_FUNCTION

FUNCTION_BLOCK T_PLC_MS_block

	VAR_OUTPUT
		T_PLC_MS :	UDINT;
	END_VAR

	VAR_EXTERNAL
		PLC_TICKS_PER_SEC :	INT;
		PLC_SYS_TICK_CNT :	DINT;
	END_VAR

	VAR
		debug :	BOOL;(*Debug-Mode ON / OFF*)
		N :	INT;(*Debug-Faktor*)
		Offset :	UDINT;(*Debug-Offset*)
		temp :	DWORD := DWORD#1;(*Debug-Offset*)
		mode :	BOOL;(*modus*)
		faktor :	UDINT;(*Systemtakt-Faktor*)
		init :	BOOL;
		v_plc_ticks_per_sec :	UDINT;
		base :	UDINT := UDINT#1000;
	END_VAR

	IF init = FALSE THEN
		v_plc_ticks_per_sec := INT_TO_UDINT(PLC_TICKS_PER_SEC);
		IF v_plc_ticks_per_sec = UDINT#1024 THEN
			faktor := UDINT#1;
			mode := FALSE;
		ELSIF v_plc_ticks_per_sec > UDINT#0 THEN
			IF v_plc_ticks_per_sec <= base THEN
				faktor := base / v_plc_ticks_per_sec;
				mode := FALSE;
			ELSE
				faktor := v_plc_ticks_per_sec / base;
				mode := TRUE;
			END_IF;
		ELSE
			faktor := UDINT#1;
		END_IF;
		init := TRUE;
	END_IF;

	IF mode THEN
		T_PLC_MS := DINT_TO_UDINT(PLC_SYS_TICK_CNT) / faktor;
	ELSE
		T_PLC_MS := DINT_TO_UDINT(PLC_SYS_TICK_CNT) * faktor;
	END_IF;

	IF debug THEN
		T_PLC_MS := (DWORD_TO_UDINT(SHL(UDINT_TO_DWORD(T_PLC_MS),N) OR SHL(temp,N)) - UDINT#1) + Offset;
	END_IF;

END_FUNCTION_BLOCK

FUNCTION_BLOCK DT_SIMU
	VAR_INPUT
		START :	UDINT;
		SPEED :	REAL := 1.0;
	END_VAR

	VAR_OUTPUT
		DTS :	UDINT;
	END_VAR

	VAR
		tc :	UDINT;
		init :	BOOL;
		last :	UDINT;
		tx :	UDINT;
		td :	UDINT;
		T_PLC_MS :	T_PLC_MS_block;
	END_VAR

	T_PLC_MS();
	tx:= T_PLC_MS.T_PLC_MS;
	tc := _REAL_TO_UDINT(UDINT_TO_REAL(tx - last) * speed);

	IF NOT init THEN
		init := TRUE;
		DTS := Start;
		tc := UDINT#0;
		last := tx;
	ELSIF SPEED = 0.0 THEN
		DTS := DTS + UDINT#1;
	ELSIF tc >= UDINT#1000 THEN
		td := (tc / UDINT#1000) * UDINT#1000;
		DTS := DTS + td;
		last := last + _REAL_TO_UDINT(UDINT_TO_REAL(td) / speed);
	END_IF;
END_FUNCTION_BLOCK

PROGRAM program0
  VAR
    LocalVar0 : UDINT;
	LocalVar1 : REAL;
	LocalOUT  : UDINT;
	func_block : DT_SIMU;
  END_VAR
	func_block.START  := LocalVar0;
	func_block.SPEED  := LocalVar1;
	func_block();
	LocalOUT := func_block.DTS;
END_PROGRAM

CONFIGURATION Config0

	VAR_GLOBAL
		PLC_TICKS_PER_SEC :	INT;
		PLC_SYS_TICK_CNT :	DINT;
	END_VAR

  	RESOURCE Res0 ON PLC
    	TASK task0(INTERVAL := T#20ms,PRIORITY := 0);
    	PROGRAM instance0 WITH task0 : program0;
  	END_RESOURCE

END_CONFIGURATION

(* ---- DT_TO_SDT.ST ---- *)
TYPE oscat_SDT :
STRUCT
	YEAR : INT;
	MONTH : INT;
	DAY : INT;
	WEEKDAY : INT;
	HOUR : INT;
	MINUTE : INT;
	SECOND : INT;
	MS : INT;
END_STRUCT;
END_TYPE

FUNCTION DT_TO_DATE2:UDINT

	VAR_INPUT
		IN :	UDINT;
	END_VAR

	DT_TO_DATE2 := (IN / UDINT#86400) * UDINT#86400;
END_FUNCTION

FUNCTION YEAR_OF_DATE:INT
	VAR_INPUT
		IDATE :	UDINT;
	END_VAR

	YEAR_OF_DATE := UDINT_TO_INT((idate+UDINT#43200) / UDINT#31557600 + UDINT#1970);
END_FUNCTION

FUNCTION DAY_OF_WEEK:INT

	VAR_INPUT
		IDATE :	UDINT;
	END_VAR

	DAY_OF_WEEK := UDINT_TO_INT((idate / UDINT#86400 + UDINT#3) MOD UDINT#7) + INT#01;
END_FUNCTION

FUNCTION LEAP_OF_DATE:BOOL

	VAR_INPUT
		IDATE :	UDINT;
	END_VAR

	LEAP_OF_DATE := SHL(UDINT_TO_DWORD((idate + UDINT#43200) / UDINT#31557600), 30) = DWORD#16#80000000;
END_FUNCTION

FUNCTION DAY_OF_YEAR:INT
	VAR_INPUT
		IDATE :	UDINT;
	END_VAR

	DAY_OF_YEAR := UDINT_TO_INT(((idate) / UDINT#86400) MOD UDINT#1461);
	IF DAY_OF_YEAR > 729 THEN
		IF DAY_OF_YEAR > 1095 THEN DAY_OF_YEAR := DAY_OF_YEAR - 1095; ELSE DAY_OF_YEAR := DAY_OF_YEAR - 729; END_IF;
	ELSIF DAY_OF_YEAR > 364 THEN
		DAY_OF_YEAR := DAY_OF_YEAR - 364;
	ELSE
		DAY_OF_YEAR := DAY_OF_YEAR + 1;
	END_IF;
END_FUNCTION

FUNCTION MONTH_OF_DATE:INT

	VAR_INPUT
		IDATE :	UDINT;
	END_VAR

	MONTH_OF_DATE := DAY_OF_YEAR(idate);
	IF MONTH_OF_DATE < 32 THEN
		MONTH_OF_DATE := 1;
	ELSIF LEAP_OF_DATE((IDATE)) THEN
		MONTH_OF_DATE := (MONTH_OF_DATE * 53 + 1668) / 1623;
	ELSE
		MONTH_OF_DATE := (MONTH_OF_DATE * 53 + 1700) / 1620;
	END_IF;
END_FUNCTION

FUNCTION DAY_OF_MONTH:INT
	VAR_INPUT
		IDATE :	UDINT;
	END_VAR

	day_of_month := day_of_year(idate);

	IF leap_of_Date((idate)) THEN
		CASE day_of_month OF
			32..60	:	day_of_month := day_of_month - 31;
			61..91	:	day_of_month := day_of_month - 60;
			92..121 :	day_of_month := day_of_month - 91;
			122..152:	day_of_month := day_of_month - 121;
			153..182:	day_of_month := day_of_month - 152;
			183..213:	day_of_month := day_of_month - 182;
			214..244:	day_of_month := day_of_month - 213;
			245..274:	day_of_month := day_of_month - 244;
			275..305:	day_of_month := day_of_month - 274;
			306..335:	day_of_month := day_of_month - 305;
			336..366:	day_of_month := day_of_month - 335;
		END_CASE;
	ELSE
		CASE day_of_month OF
			32..59	:	day_of_month := day_of_month - 31;
			60..90	:	day_of_month := day_of_month - 59;
			91..120 :	day_of_month := day_of_month - 90;
			121..151:	day_of_month := day_of_month - 120;
			152..181:	day_of_month := day_of_month - 151;
			182..212:	day_of_month := day_of_month - 181;
			213..243:	day_of_month := day_of_month - 212;
			244..273:	day_of_month := day_of_month - 243;
			274..304:	day_of_month := day_of_month - 273;
			305..334:	day_of_month := day_of_month - 304;
			335..365:	day_of_month := day_of_month - 334;
		END_CASE;
	END_IF;
END_FUNCTION

FUNCTION _INT_TO_UDINT:UDINT
	VAR_INPUT
		IN :	INT;
	END_VAR

	_INT_TO_UDINT := DINT_TO_UDINT(INT_TO_DINT(IN));
END_FUNCTION

FUNCTION_BLOCK DT_TO_SDT

	VAR_INPUT
		DTI :	UDINT;
	END_VAR

	VAR_OUTPUT
		SDT :	oscat_SDT;
	END_VAR

	VAR
		tmp :	UDINT;
		tdt :	UDINT;
	END_VAR

	tmp := DT_TO_DATE2(dti);
	tdt := dti - tmp;
	SDT.YEAR := YEAR_OF_DATE(tmp);
	SDT.MONTH := MONTH_OF_DATE(tmp);
	SDT.DAY := DAY_OF_MONTH(tmp);
	SDT.WEEKDAY := DAY_OF_WEEK(tmp);
	SDT.SECOND := UDINT_TO_INT(tdt MOD UDINT#60);
	SDT.MINUTE := UDINT_TO_INT((tdt / UDINT#60) MOD UDINT#60);
	SDT.HOUR := UDINT_TO_INT(tdt / UDINT#3600);

END_FUNCTION_BLOCK

PROGRAM program0
  VAR
    LocalVar0 : UDINT;
	LocalOUT  : oscat_SDT;
	func_block : DT_TO_SDT;
  END_VAR
	func_block.DTI  := LocalVar0;
	func_block();
	LocalOUT := func_block.SDT;
END_PROGRAM

CONFIGURATION Config0
  RESOURCE Res0 ON PLC
    TASK task0(INTERVAL := T#20ms,PRIORITY := 0);
    PROGRAM instance0 WITH task0 : program0;
  END_RESOURCE
END_CONFIGURATION

(* ---- DT_TO_STRING.ST ---- *)
FUNCTION YEAR_OF_DATE:INT
	VAR_INPUT
		IDATE :	UDINT;
	END_VAR

	YEAR_OF_DATE := UDINT_TO_INT((idate+UDINT#43200) / UDINT#31557600 + UDINT#1970);
END_FUNCTION

FUNCTION DAY_OF_YEAR:INT
	VAR_INPUT
		IDATE :	UDINT;
	END_VAR

	DAY_OF_YEAR := UDINT_TO_INT(((idate) / UDINT#86400) MOD UDINT#1461);
	IF DAY_OF_YEAR > 729 THEN
		IF DAY_OF_YEAR > 1095 THEN DAY_OF_YEAR := DAY_OF_YEAR - 1095; ELSE DAY_OF_YEAR := DAY_OF_YEAR - 729; END_IF;
	ELSIF DAY_OF_YEAR > 364 THEN
		DAY_OF_YEAR := DAY_OF_YEAR - 364;
	ELSE
		DAY_OF_YEAR := DAY_OF_YEAR + 1;
	END_IF;
END_FUNCTION

FUNCTION LEAP_OF_DATE:BOOL

	VAR_INPUT
		IDATE :	UDINT;
	END_VAR

	LEAP_OF_DATE := SHL(UDINT_TO_DWORD((idate + UDINT#43200) / UDINT#31557600), 30) = DWORD#16#80000000;
END_FUNCTION

FUNCTION MONTH_OF_DATE:INT

	VAR_INPUT
		IDATE :	UDINT;
	END_VAR

	MONTH_OF_DATE := DAY_OF_YEAR(idate);
	IF MONTH_OF_DATE < 32 THEN
		MONTH_OF_DATE := 1;
	ELSIF LEAP_OF_DATE(IDATE) THEN
		MONTH_OF_DATE := (MONTH_OF_DATE * 53 + 1668) / 1623;
	ELSE
		MONTH_OF_DATE := (MONTH_OF_DATE * 53 + 1700) / 1620;
	END_IF;
END_FUNCTION

FUNCTION DAY_OF_MONTH:INT
	VAR_INPUT
		IDATE :	UDINT;
	END_VAR

	day_of_month := day_of_year(idate);

	IF leap_of_Date((idate)) THEN
		CASE day_of_month OF
			32..60	:	day_of_month := day_of_month - 31;
			61..91	:	day_of_month := day_of_month - 60;
			92..121 :	day_of_month := day_of_month - 91;
			122..152:	day_of_month := day_of_month - 121;
			153..182:	day_of_month := day_of_month - 152;
			183..213:	day_of_month := day_of_month - 182;
			214..244:	day_of_month := day_of_month - 213;
			245..274:	day_of_month := day_of_month - 244;
			275..305:	day_of_month := day_of_month - 274;
			306..335:	day_of_month := day_of_month - 305;
			336..366:	day_of_month := day_of_month - 335;
		END_CASE;
	ELSE
		CASE day_of_month OF
			32..59	:	day_of_month := day_of_month - 31;
			60..90	:	day_of_month := day_of_month - 59;
			91..120 :	day_of_month := day_of_month - 90;
			121..151:	day_of_month := day_of_month - 120;
			152..181:	day_of_month := day_of_month - 151;
			182..212:	day_of_month := day_of_month - 181;
			213..243:	day_of_month := day_of_month - 212;
			244..273:	day_of_month := day_of_month - 243;
			274..304:	day_of_month := day_of_month - 273;
			305..334:	day_of_month := day_of_month - 304;
			335..365:	day_of_month := day_of_month - 334;
		END_CASE;
	END_IF;
END_FUNCTION

FUNCTION SECOND_OF_DT:INT

	VAR_INPUT
		XDT :	UDINT;
	END_VAR

	SECOND_OF_DT := UDINT_TO_INT(XDT MOD UDINT#60);
END_FUNCTION

FUNCTION HOUR_OF_DT:INT
	VAR_INPUT
		XDT :	UDINT;
	END_VAR

	HOUR_OF_DT := UDINT_TO_INT((XDT MOD UDINT#86400) / UDINT#3600);
END_FUNCTION

FUNCTION MINUTE_OF_DT:INT
	VAR_INPUT
		XDT :	UDINT;
	END_VAR

	MINUTE_OF_DT := UDINT_TO_INT((XDT MOD UDINT#3600) / UDINT#60);
END_FUNCTION

FUNCTION_BLOCK DT_TO_STRING_Block

	VAR_INPUT
		IDT :	UDINT;
	END_VAR

	VAR_OUTPUT
		DT_STRING :	STRING;
	END_VAR

	VAR
		st_tmp1 :	STRING;
		st_tmp2 :	STRING;
	END_VAR

	st_tmp2 := CONCAT(INT_TO_STRING(YEAR_OF_DATE(IDT)),INT_TO_STRING(MONTH_OF_DATE(IDT)));
	st_tmp1 := CONCAT(INT_TO_STRING(day_of_month(IDT)),INT_TO_STRING(hour_of_DT(IDT)));
	st_tmp2 := CONCAT(st_tmp2,st_tmp1);
	st_tmp1 := CONCAT(INT_TO_STRING(minute_of_DT(IDT)),INT_TO_STRING(second_of_DT(IDT)));
	st_tmp2 := CONCAT(st_tmp2,st_tmp1);
	DT_STRING := st_tmp2;
END_FUNCTION_BLOCK

PROGRAM program0
	VAR
		IDT : UDINT;
		OUT  : STRING;
		func_block : DT_TO_STRING_Block;
	END_VAR
	func_block.IDT := IDT;
	func_block();
	OUT := func_block.DT_STRING;
END_PROGRAM

CONFIGURATION Config0
	RESOURCE Res0 ON PLC
		TASK task0(INTERVAL := T#20ms,PRIORITY := 0);
		PROGRAM instance0 WITH task0 : program0;
	END_RESOURCE
END_CONFIGURATION

(* ---- DWORD_TO_STRB.ST ---- *)
FUNCTION_BLOCK DWORD_TO_STRB_Block
	VAR_INPUT
		IN :	DWORD;
	END_VAR

	VAR_OUTPUT
		DWORD_TO_STRB :	STRING;
	END_VAR

	VAR
		i :	INT;
	END_VAR

	DWORD_TO_STRB :='';
	FOR i := 1 TO 32 DO
		IF (in AND DWORD#16#8000_0000) > DWORD#0 THEN
			DWORD_TO_STRB := CONCAT(DWORD_TO_STRB,'1');
		ELSE
			DWORD_TO_STRB := CONCAT(DWORD_TO_STRB,'0');
		END_IF;
		in := SHL(in, 1);
	END_FOR;
END_FUNCTION_BLOCK

PROGRAM program0
  VAR
    IN :	DWORD;

	DWORD_TO_STRB :	STRING;
	func_block : DWORD_TO_STRB_Block;
  END_VAR
	func_block.IN  := IN;
	func_block();
	DWORD_TO_STRB := func_block.DWORD_TO_STRB;
END_PROGRAM

CONFIGURATION Config0
  RESOURCE Res0 ON PLC
    TASK task0(INTERVAL := T#20ms,PRIORITY := 0);
    PROGRAM instance0 WITH task0 : program0;
  END_RESOURCE
END_CONFIGURATION

(* ---- DWORD_TO_STRF.ST ---- *)
FUNCTION_BLOCK DWORD_TO_STRF_Block

	VAR_INPUT
		IN :	DWORD;
		N :	INT;
	END_VAR

	VAR_OUTPUT
		DWORD_TO_STRF :	STRING;
	END_VAR

	VAR
		temp :	STRING;
		temp2 :	STRING;
		L : INT;
	END_VAR

	temp := DWORD_TO_STRING(in);
	L := LEN(temp);
	IF N < L THEN
		temp :=RIGHT(temp,N);
		L := N;
	END_IF;

	WHILE L < N DO
		temp2 := temp;
		temp := CONCAT('0', temp2);
		L := L + 1;
	END_WHILE;
	DWORD_TO_STRF := temp;

END_FUNCTION_BLOCK

PROGRAM program0
  VAR
    IN :	DWORD;
	N :		INT;
	DWORD_TO_STRF :	STRING;
	func_block : DWORD_TO_STRF_Block;
  END_VAR
	func_block.IN  := IN;
	func_block.N  := N;
	func_block();
	DWORD_TO_STRF := func_block.DWORD_TO_STRF;
END_PROGRAM

CONFIGURATION Config0
  RESOURCE Res0 ON PLC
    TASK task0(INTERVAL := T#20ms,PRIORITY := 0);
    PROGRAM instance0 WITH task0 : program0;
  END_RESOURCE
END_CONFIGURATION

(* ---- DWORD_TO_STRH.ST ---- *)
FUNCTION_BLOCK DWORD_TO_STRH_Block

	VAR_INPUT
		IN :	DWORD;
	END_VAR

	VAR_OUTPUT
		DWORD_TO_STRH :	STRING;
	END_VAR

	DWORD_TO_STRH:=DWORD_TO_STRING(IN);

END_FUNCTION_BLOCK

PROGRAM program0
  VAR
    LocalVar0 : DWORD;
	LocalOUT  : STRING;
	func_block : DWORD_TO_STRH_Block;
  END_VAR
	func_block.IN  := LocalVar0;
	func_block();
	LocalOUT := func_block.DWORD_TO_STRH;
END_PROGRAM

CONFIGURATION Config0
  RESOURCE Res0 ON PLC
    TASK task0(INTERVAL := T#20ms,PRIORITY := 0);
    PROGRAM instance0 WITH task0 : program0;
  END_RESOURCE
END_CONFIGURATION

(* ---- ENERGY.ST ---- *)
FUNCTION_BLOCK ENERGY
	VAR_INPUT
		J :	REAL;
		C :	REAL;
		WH :	REAL;
	END_VAR

	VAR_OUTPUT
		YJ :	REAL;
		YC :	REAL;
		YWH :	REAL;
	END_VAR

	YJ := J + Wh * 3600.0 + C * 4.1868;
	YC := YJ * 0.238845896627496;
	YWh := YJ * 2.7777777778E-004;
END_FUNCTION_BLOCK

PROGRAM program0
  VAR
		J  :	REAL;
		C  :	REAL;
		WH :	REAL;

		YJ  :	REAL;
		YC  :	REAL;
		YWH :	REAL;
	func_block : ENERGY;
  END_VAR
	func_block.J  :=J ;
	func_block.C  :=C ;
	func_block.WH :=WH;
	func_block();
	YJ  := func_block.YJ ;
	YC  := func_block.YC ;
	YWH := func_block.YWH;

END_PROGRAM

CONFIGURATION Config0
	RESOURCE Res0 ON PLC
		TASK task0(INTERVAL := T#20ms,PRIORITY := 0);
		PROGRAM instance0 WITH task0 : program0;
	END_RESOURCE
END_CONFIGURATION

(* ---- ESR_COLLECT.ST ---- *)
TYPE
	oscat_esr_collect_data      : ARRAY [0..7]    OF BYTE;
END_TYPE
TYPE oscat_esr_data :
  STRUCT
	typ    : BYTE;
	adress : STRING;
	DS     : UDINT;
	TS     : TIME;
	data   : oscat_esr_collect_data;
  END_STRUCT;
END_TYPE

TYPE
  oscat_ESR_3                : ARRAY [0..3] OF oscat_esr_data;
  oscat_ESR_31               : ARRAY [0..31] OF oscat_esr_data;
END_TYPE

FUNCTION INC1:INT

	VAR_INPUT
		X :	INT;
		N :	INT;
	END_VAR

	IF X >= N - 1 THEN
		INC1 := 0;
	ELSE
		INC1 := X + 1;
	END_IF;
END_FUNCTION

FUNCTION_BLOCK ESR_COLLECT
	VAR_INPUT
		ESR_0 :	oscat_ESR_3;
		ESR_1 :	oscat_ESR_3;
		ESR_2 :	oscat_ESR_3;
		ESR_3 :	oscat_ESR_3;
		ESR_4 :	oscat_ESR_3;
		ESR_5 :	oscat_ESR_3;
		ESR_6 :	oscat_ESR_3;
		ESR_7 :	oscat_ESR_3;
		RST :	BOOL;
	END_VAR

	VAR_IN_OUT
		POS :	INT;
	END_VAR

	VAR_OUTPUT
		ESR_OUT :	oscat_ESR_31;
	END_VAR

	VAR
		cnt :	INT := -1;
		max_in :	INT := 3;
		max_out :	INT := 32;
	END_VAR

	IF rst OR cnt < 0 THEN
		pos := -1;
	ELSE
		FOR cnt := 0 TO max_in DO
		IF esr_0[cnt].typ > BYTE#0 THEN pos := INC1(pos, max_out); esr_out[pos] := esr_0[cnt]; END_IF;
		IF esr_1[cnt].typ > BYTE#0 THEN pos := INC1(pos, max_out); esr_out[pos] := esr_1[cnt]; END_IF;
		IF esr_2[cnt].typ > BYTE#0 THEN pos := INC1(pos, max_out); esr_out[pos] := esr_2[cnt]; END_IF;
		IF esr_3[cnt].typ > BYTE#0 THEN pos := INC1(pos, max_out); esr_out[pos] := esr_3[cnt]; END_IF;
		IF esr_4[cnt].typ > BYTE#0 THEN pos := INC1(pos, max_out); esr_out[pos] := esr_4[cnt]; END_IF;
		IF esr_5[cnt].typ > BYTE#0 THEN pos := INC1(pos, max_out); esr_out[pos] := esr_5[cnt]; END_IF;
		IF esr_6[cnt].typ > BYTE#0 THEN pos := INC1(pos, max_out); esr_out[pos] := esr_6[cnt]; END_IF;
		IF esr_7[cnt].typ > BYTE#0 THEN pos := INC1(pos, max_out); esr_out[pos] := esr_7[cnt]; END_IF;
	END_FOR;
	END_IF;

END_FUNCTION_BLOCK

PROGRAM program0
  VAR
	ESR_0 :	oscat_ESR_3;
	ESR_1 :	oscat_ESR_3;
	ESR_2 :	oscat_ESR_3;
	ESR_3 :	oscat_ESR_3;
	ESR_4 :	oscat_ESR_3;
	ESR_5 :	oscat_ESR_3;
	ESR_6 :	oscat_ESR_3;
	ESR_7 :	oscat_ESR_3;
	RST   :	BOOL;

	POS   :	INT;

	ESR_OUT :	oscat_ESR_31;

	func_block : ESR_COLLECT;
  END_VAR
	func_block.ESR_0 :=ESR_0;
	func_block.ESR_1 :=ESR_1;
	func_block.ESR_2 :=ESR_2;
	func_block.ESR_3 :=ESR_3;
	func_block.ESR_4 :=ESR_4;
	func_block.ESR_5 :=ESR_5;
	func_block.ESR_6 :=ESR_6;
	func_block.ESR_7 :=ESR_7;
	func_block.RST   :=RST  ;
	func_block.POS   :=POS  ;

	func_block();
	POS := func_block.POS;
	ESR_OUT := func_block.ESR_OUT;

END_PROGRAM

CONFIGURATION Config0
	RESOURCE Res0 ON PLC
		TASK task0(INTERVAL := T#20ms,PRIORITY := 0);
		PROGRAM instance0 WITH task0 : program0;
	END_RESOURCE
END_CONFIGURATION

(* ---- ESR_MON_B8.ST ---- *)
TYPE
	oscat_esr_collect_data      : ARRAY [0..7]    OF BYTE;
END_TYPE
TYPE oscat_esr_data :
  STRUCT
	typ    : BYTE;
	adress : STRING;
	DS     : UDINT;
	TS     : TIME;
	data   : oscat_esr_collect_data;
  END_STRUCT;
END_TYPE

TYPE
  oscat_ESR_3                : ARRAY [0..3] OF oscat_esr_data;
  oscat_ESR_31               : ARRAY [0..31] OF oscat_esr_data;
END_TYPE

FUNCTION_BLOCK T_PLC_MS_block

	VAR_OUTPUT
		T_PLC_MS :	UDINT;
	END_VAR

	VAR_EXTERNAL
		PLC_TICKS_PER_SEC :	INT;
		PLC_SYS_TICK_CNT :	DINT;
	END_VAR

	VAR
		debug :	BOOL;(*Debug-Mode ON / OFF*)
		N :	INT;(*Debug-Faktor*)
		Offset :	UDINT;(*Debug-Offset*)
		temp :	DWORD := DWORD#1;(*Debug-Offset*)
		mode :	BOOL;(*modus*)
		faktor :	UDINT;(*Systemtakt-Faktor*)
		init :	BOOL;
		v_plc_ticks_per_sec :	UDINT;
		base :	UDINT := UDINT#1000;
	END_VAR

	IF init = FALSE THEN
		v_plc_ticks_per_sec := INT_TO_UDINT(PLC_TICKS_PER_SEC);
		IF v_plc_ticks_per_sec = UDINT#1024 THEN
			faktor := UDINT#1;
			mode := FALSE;
		ELSIF v_plc_ticks_per_sec > UDINT#0 THEN
			IF v_plc_ticks_per_sec <= base THEN
				faktor := base / v_plc_ticks_per_sec;
				mode := FALSE;
			ELSE
				faktor := v_plc_ticks_per_sec / base;
				mode := TRUE;
			END_IF;
		ELSE
			faktor := UDINT#1;
		END_IF;
		init := TRUE;
	END_IF;

	IF mode THEN
		T_PLC_MS := DINT_TO_UDINT(PLC_SYS_TICK_CNT) / faktor;
	ELSE
		T_PLC_MS := DINT_TO_UDINT(PLC_SYS_TICK_CNT) * faktor;
	END_IF;

	IF debug THEN
		T_PLC_MS := (DWORD_TO_UDINT(SHL(UDINT_TO_DWORD(T_PLC_MS),N) OR SHL(temp,N)) - UDINT#1) + Offset;
	END_IF;

END_FUNCTION_BLOCK

FUNCTION_BLOCK ESR_MON_B8

	VAR_INPUT
		S0 :	BOOL;
		A0 :	STRING;
		S1 :	BOOL;
		A1 :	STRING;
		S2 :	BOOL;
		A2 :	STRING;
		S3 :	BOOL;
		A3 :	STRING;
		S4 :	BOOL;
		A4 :	STRING;
		S5 :	BOOL;
		A5 :	STRING;
		S6 :	BOOL;
		A6 :	STRING;
		S7 :	BOOL;
		A7 :	STRING;
		DT_IN :	UDINT;
	END_VAR

	VAR_IN_OUT
		ESR_Out :	oscat_ESR_3;
	END_VAR

	VAR_OUTPUT
		ESR_FLAG :	BOOL;
	END_VAR

	VAR
		x0 :	BOOL;
		x1 :	BOOL;
		x2 :	BOOL;
		x3 :	BOOL;
		x4 :	BOOL;
		x5 :	BOOL;
		x6 :	BOOL;
		x7 :	BOOL;
		tx :	TIME;
		cnt :	INT;
		T_PLC_MS :	T_PLC_MS_block;
	END_VAR

	T_PLC_MS();
	tx:= UDINT_TO_TIME(T_PLC_MS.T_PLC_MS);

	ESR_Flag := FALSE;
	esr_out[3].typ := BYTE#0;
	esr_out[2].typ := BYTE#0;
	esr_out[1].typ := BYTE#0;
	esr_out[0].typ := BYTE#0;
	cnt := 0;

	IF s0 <> X0 THEN
		esr_out[cnt].typ := INT_TO_BYTE(10 + BOOL_TO_INT(s0));
		esr_out[cnt].adress := a0;
		esr_out[cnt].DS := DT_in;
		esr_out[cnt].TS := TX;
		X0 := S0;
		cnt := cnt + 1;
		esr_flag := TRUE;
	END_IF;
	IF s1 <> X1 THEN
		esr_out[cnt].typ := INT_TO_BYTE(10 + BOOL_TO_INT(s1));
		esr_out[cnt].adress := a1;
		esr_out[cnt].DS := DT_in;
		esr_out[cnt].TS := TX;
		X1 := S1;
		cnt := cnt + 1;
		esr_flag := TRUE;
	END_IF;
	IF s2 <> X2 THEN
		esr_out[cnt].typ := INT_TO_BYTE(10 + BOOL_TO_INT(s2));
		esr_out[cnt].adress := a2;
		esr_out[cnt].DS := DT_in;
		esr_out[cnt].TS := TX;
		X2 := S2;
		cnt := cnt + 1;
		esr_flag := TRUE;
	END_IF;
	IF s3 <> X3 THEN
		esr_out[cnt].typ := INT_TO_BYTE(10 + BOOL_TO_INT(s3));
		esr_out[cnt].adress := a3;
		esr_out[cnt].DS := DT_in;
		esr_out[cnt].TS := TX;
		X3 := S3;
		cnt := cnt + 1;
		esr_flag := TRUE;
	END_IF;
	IF s4 <> X4 AND cnt < 4 THEN
		esr_out[cnt].typ := INT_TO_BYTE(10 + BOOL_TO_INT(s4));
		esr_out[cnt].adress := a4;
		esr_out[cnt].DS := DT_in;
		esr_out[cnt].TS := TX;
		X4 := S4;
		cnt := cnt + 1;
		esr_flag := TRUE;
	END_IF;
	IF s5 <> X5  AND cnt < 4 THEN
		esr_out[cnt].typ := INT_TO_BYTE(10 + BOOL_TO_INT(s5));
		esr_out[cnt].adress := a5;
		esr_out[cnt].DS := DT_in;
		esr_out[cnt].TS := TX;
		X5 := S5;
		cnt := cnt + 1;
		esr_flag := TRUE;
	END_IF;
	IF s6 <> X6  AND cnt < 4 THEN
		esr_out[cnt].typ := INT_TO_BYTE(10 + BOOL_TO_INT(s6));
		esr_out[cnt].adress := a6;
		esr_out[cnt].DS := DT_in;
		esr_out[cnt].TS := TX;
		X6 := S6;
		cnt := cnt + 1;
		esr_flag := TRUE;
	END_IF;
	IF s7 <> X7  AND cnt < 4 THEN
		esr_out[cnt].typ := INT_TO_BYTE(10 + BOOL_TO_INT(s7));
		esr_out[cnt].adress := a7;
		esr_out[cnt].DS := DT_in;
		esr_out[cnt].TS := TX;
		X7 := S7;
		cnt := cnt + 1;
		esr_flag := TRUE;
	END_IF;

END_FUNCTION_BLOCK

PROGRAM program0

	VAR

		S0 :	BOOL;
		A0 :	STRING;
		S1 :	BOOL;
		A1 :	STRING;
		S2 :	BOOL;
		A2 :	STRING;
		S3 :	BOOL;
		A3 :	STRING;
		S4 :	BOOL;
		A4 :	STRING;
		S5 :	BOOL;
		A5 :	STRING;
		S6 :	BOOL;
		A6 :	STRING;
		S7 :	BOOL;
		A7 :	STRING;
		DT_IN   :	UDINT;

		ESR_Out :	oscat_ESR_3;

		ESR_FLAG :	BOOL;

		func_block : ESR_MON_B8;
  	END_VAR
	func_block.S0 := S0;
	func_block.A0 := A0;
	func_block.S1 := S1;
	func_block.A1 := A1;
	func_block.S2 := S2;
	func_block.A2 := A2;
	func_block.S3 := S3;
	func_block.A3 := A3;
	func_block.S4 := S4;
	func_block.A4 := A4;
	func_block.S5 := S5;
	func_block.A5 := A5;
	func_block.S6 := S6;
	func_block.A6 := A6;
	func_block.S7 := S7;
	func_block.A7 := A7;
	func_block.DT_IN := DT_IN;
	func_block.ESR_Out := ESR_Out;
	func_block();
	ESR_Out := func_block.ESR_Out;
	ESR_FLAG := func_block.ESR_FLAG;

END_PROGRAM

CONFIGURATION Config0

	VAR_GLOBAL
		PLC_TICKS_PER_SEC :	INT;
		PLC_SYS_TICK_CNT :	DINT;
	END_VAR

  	RESOURCE Res0 ON PLC
    	TASK task0(INTERVAL := T#20ms,PRIORITY := 0);
    	PROGRAM instance0 WITH task0 : program0;
  	END_RESOURCE

END_CONFIGURATION

(* ---- ESR_MON_X8.ST ---- *)
TYPE
	oscat_esr_collect_data      : ARRAY [0..7]    OF BYTE;
END_TYPE

TYPE oscat_esr_data :
  STRUCT
	typ    : BYTE;
	adress : STRING;
	DS     : UDINT;
	TS     : TIME;
	data   : oscat_esr_collect_data;
  END_STRUCT;
END_TYPE

TYPE
  oscat_ESR_3                : ARRAY [0..3] OF oscat_esr_data;
  oscat_ESR_31               : ARRAY [0..31] OF oscat_esr_data;
END_TYPE

FUNCTION_BLOCK STATUS_TO_ESR_Block

	VAR_INPUT
		STATUS :	BYTE;
		ADRESS :	STRING;
		DT_IN :	UDINT;
		TS :	TIME;
	END_VAR

	VAR_OUTPUT
		STATUS_TO_ESR :	oscat_esr_data;
	END_VAR

	IF status < BYTE#100 THEN
		status_to_ESR.typ := BYTE#1;
	ELSIF status < BYTE#200 THEN
		status_to_ESR.typ := BYTE#2;
	ELSE
		status_to_ESR.typ := BYTE#3;
	END_IF;
	status_to_ESR.adress:= adress;
	status_to_ESR.DS := DT_in;
	status_to_ESR.TS := TS;
	status_to_ESR.data[0] := status;
END_FUNCTION_BLOCK

FUNCTION_BLOCK T_PLC_MS_block

	VAR_OUTPUT
		T_PLC_MS :	UDINT;
	END_VAR

	VAR_EXTERNAL
		PLC_TICKS_PER_SEC :	INT;
		PLC_SYS_TICK_CNT :	DINT;
	END_VAR

	VAR
		debug :	BOOL;(*Debug-Mode ON / OFF*)
		N :	INT;(*Debug-Faktor*)
		Offset :	UDINT;(*Debug-Offset*)
		temp :	DWORD := DWORD#1;(*Debug-Offset*)
		mode :	BOOL;(*modus*)
		faktor :	UDINT;(*Systemtakt-Faktor*)
		init :	BOOL;
		v_plc_ticks_per_sec :	UDINT;
		base :	UDINT := UDINT#1000;
	END_VAR

	IF init = FALSE THEN
		v_plc_ticks_per_sec := INT_TO_UDINT(PLC_TICKS_PER_SEC);
		IF v_plc_ticks_per_sec = UDINT#1024 THEN
			faktor := UDINT#1;
			mode := FALSE;
		ELSIF v_plc_ticks_per_sec > UDINT#0 THEN
			IF v_plc_ticks_per_sec <= base THEN
				faktor := base / v_plc_ticks_per_sec;
				mode := FALSE;
			ELSE
				faktor := v_plc_ticks_per_sec / base;
				mode := TRUE;
			END_IF;
		ELSE
			faktor := UDINT#1;
		END_IF;
		init := TRUE;
	END_IF;

	IF mode THEN
		T_PLC_MS := DINT_TO_UDINT(PLC_SYS_TICK_CNT) / faktor;
	ELSE
		T_PLC_MS := DINT_TO_UDINT(PLC_SYS_TICK_CNT) * faktor;
	END_IF;

	IF debug THEN
		T_PLC_MS := (DWORD_TO_UDINT(SHL(UDINT_TO_DWORD(T_PLC_MS),N) OR SHL(temp,N)) - UDINT#1) + Offset;
	END_IF;

END_FUNCTION_BLOCK

FUNCTION_BLOCK ESR_MON_X8
	VAR_INPUT
		S0 :	BYTE;
		A0 :	STRING;
		S1 :	BYTE;
		A1 :	STRING;
		S2 :	BYTE;
		A2 :	STRING;
		S3 :	BYTE;
		A3 :	STRING;
		S4 :	BYTE;
		A4 :	STRING;
		S5 :	BYTE;
		A5 :	STRING;
		S6 :	BYTE;
		A6 :	STRING;
		S7 :	BYTE;
		A7 :	STRING;
		DT_IN :	UDINT;
		MODE :	BYTE := BYTE#3;
	END_VAR

	VAR_IN_OUT
		ESR_OUT :	oscat_ESR_3;
	END_VAR

	VAR_OUTPUT
		ESR_FLAG :	BOOL;
	END_VAR

	VAR
		x0 :	BYTE;
		x1 :	BYTE;
		x2 :	BYTE;
		x3 :	BYTE;
		x4 :	BYTE;
		x5 :	BYTE;
		x6 :	BYTE;
		x7 :	BYTE;
		tx :	TIME;
		cnt :	INT;
		status_to_ESR :	STATUS_TO_ESR_Block;
		T_PLC_MS :	T_PLC_MS_block;
	END_VAR

	T_PLC_MS();
	tx:= UDINT_TO_TIME(T_PLC_MS.T_PLC_MS);

	ESR_Flag := FALSE;
	esr_out[3].typ := BYTE#0;
	esr_out[2].typ := BYTE#0;
	esr_out[1].typ := BYTE#0;
	esr_out[0].typ := BYTE#0;
	cnt := 0;

	IF s0 <> X0 AND ((s0 < BYTE#100) OR (S0 > BYTE#99 AND S0 < BYTE#200 AND mode >= BYTE#2) OR (S0 > BYTE#199 AND mode = BYTE#3)) THEN

		status_to_ESR.status := s0;
		status_to_ESR.adress := a0;
		status_to_ESR.DT_in  := DT_in;
		status_to_ESR.TS     := tx;
		status_to_ESR();
		esr_out[cnt] := status_to_ESR.status_to_ESR;

		X0 := S0;
		cnt := cnt + 1;
		esr_flag := TRUE;
	END_IF;
	IF s1 <> X1 AND ((s1 < BYTE#100) OR (S1 > BYTE#99 AND S1 < BYTE#200 AND mode >= BYTE#2) OR (S1 > BYTE#199 AND mode = BYTE#3)) THEN

		status_to_ESR.status := s1;
		status_to_ESR.adress := a1;
		status_to_ESR.DT_in  := DT_in;
		status_to_ESR.TS     := tx;
		status_to_ESR();
		esr_out[cnt] := status_to_ESR.status_to_ESR;

		X1 := S1;
		cnt := cnt + 1;
		esr_flag := TRUE;
	END_IF;
	IF s2 <> X2 AND ((s2 < BYTE#100) OR (S2 > BYTE#99 AND S2 < BYTE#200 AND mode >= BYTE#2) OR (S2 > BYTE#199 AND mode = BYTE#3)) THEN

		status_to_ESR.status := s2;
		status_to_ESR.adress := a2;
		status_to_ESR.DT_in  := DT_in;
		status_to_ESR.TS     := tx;
		status_to_ESR();
		esr_out[cnt] := status_to_ESR.status_to_ESR;

		X2 := S2;
		cnt := cnt + 1;
		esr_flag := TRUE;
	END_IF;
	IF s3 <> X3 AND ((s3 < BYTE#100) OR (S3 > BYTE#99 AND S3 < BYTE#200 AND mode >= BYTE#2) OR (S3 > BYTE#199 AND mode = BYTE#3)) THEN

		status_to_ESR.status := s3;
		status_to_ESR.adress := a3;
		status_to_ESR.DT_in  := DT_in;
		status_to_ESR.TS     := tx;
		status_to_ESR();
		esr_out[cnt] := status_to_ESR.status_to_ESR;

		X3 := S3;
		cnt := cnt + 1;
		esr_flag := TRUE;
	END_IF;
	IF cnt < 4 AND s4 <> X4 AND ((s4 < BYTE#100) OR (S4 > BYTE#99 AND S4 < BYTE#200 AND mode >= BYTE#2) OR (S4 > BYTE#199 AND mode = BYTE#3)) THEN

		status_to_ESR.status := s4;
		status_to_ESR.adress := a4;
		status_to_ESR.DT_in  := DT_in;
		status_to_ESR.TS     := tx;
		status_to_ESR();
		esr_out[cnt] := status_to_ESR.status_to_ESR;

		X4 := S4;
		cnt := cnt + 1;
		esr_flag := TRUE;
	END_IF;
	IF cnt < 4 AND s5 <> X5 AND ((s5 < BYTE#100) OR (S5 > BYTE#99 AND S5 < BYTE#200 AND mode >= BYTE#2) OR (S5 > BYTE#199 AND mode = BYTE#3)) THEN

		status_to_ESR.status := s5;
		status_to_ESR.adress := a5;
		status_to_ESR.DT_in  := DT_in;
		status_to_ESR.TS     := tx;
		status_to_ESR();
		esr_out[cnt] := status_to_ESR.status_to_ESR;

		X5 := S5;
		cnt := cnt + 1;
		esr_flag := TRUE;
	END_IF;
	IF cnt < 4 AND s6 <> X6 AND ((s6 < BYTE#100) OR (S6 > BYTE#99 AND S6 < BYTE#200 AND mode >= BYTE#2) OR (S6 > BYTE#199 AND mode = BYTE#3)) THEN

		status_to_ESR.status := s6;
		status_to_ESR.adress := a6;
		status_to_ESR.DT_in  := DT_in;
		status_to_ESR.TS     := tx;
		status_to_ESR();
		esr_out[cnt] := status_to_ESR.status_to_ESR;

		X6 := S6;
		cnt := cnt + 1;
		esr_flag := TRUE;
	END_IF;
	IF cnt < 4 AND s7 <> X7 AND ((s7 < BYTE#100) OR (S7 > BYTE#99 AND S7 < BYTE#200 AND mode >= BYTE#2) OR (S7 > BYTE#199 AND mode = BYTE#3)) THEN

		status_to_ESR.status := s7;
		status_to_ESR.adress := a7;
		status_to_ESR.DT_in  := DT_in;
		status_to_ESR.TS     := tx;
		status_to_ESR();
		esr_out[cnt] := status_to_ESR.status_to_ESR;

		X7 := S7;
		cnt := cnt + 1;
		esr_flag := TRUE;
	END_IF;

END_FUNCTION_BLOCK

PROGRAM program0

	VAR
	S0 :	BYTE;
	A0 :	STRING;
	S1 :	BYTE;
	A1 :	STRING;
	S2 :	BYTE;
	A2 :	STRING;
	S3 :	BYTE;
	A3 :	STRING;
	S4 :	BYTE;
	A4 :	STRING;
	S5 :	BYTE;
	A5 :	STRING;
	S6 :	BYTE;
	A6 :	STRING;
	S7 :	BYTE;
	A7 :	STRING;
	DT_IN :	UDINT;
	MODE :	BYTE;

	ESR_OUT :	oscat_ESR_3;

	ESR_FLAG :	BOOL;

		func_block : ESR_MON_X8;
  	END_VAR
	func_block.S0 := S0;
	func_block.A0 := A0;
	func_block.S1 := S1;
	func_block.A1 := A1;
	func_block.S2 := S2;
	func_block.A2 := A2;
	func_block.S3 := S3;
	func_block.A3 := A3;
	func_block.S4 := S4;
	func_block.A4 := A4;
	func_block.S5 := S5;
	func_block.A5 := A5;
	func_block.S6 := S6;
	func_block.A6 := A6;
	func_block.S7 := S7;
	func_block.A7 := A7;
	func_block.DT_IN := DT_IN;
	func_block.MODE := MODE;
	func_block.ESR_Out := ESR_Out;
	func_block();
	ESR_Out := func_block.ESR_Out;
	ESR_FLAG := func_block.ESR_FLAG;
END_PROGRAM

CONFIGURATION Config0

	VAR_GLOBAL
		PLC_TICKS_PER_SEC :	INT;
		PLC_SYS_TICK_CNT :	DINT;
	END_VAR

  	RESOURCE Res0 ON PLC
    	TASK task0(INTERVAL := T#20ms,PRIORITY := 0);
    	PROGRAM instance0 WITH task0 : program0;
  	END_RESOURCE

END_CONFIGURATION

(* ---- EVENTS.ST ---- *)
TYPE oscat_HOLIDAY_DATA :
  STRUCT
	NAME : STRING;
	DAY : SINT;
	MONTH : SINT;
	USE : SINT;
	PAD_BYTE : BYTE;
  END_STRUCT;
END_TYPE

TYPE
  oscat_HOLIDAY_DATA_0_29 	: ARRAY [0..29] OF oscat_HOLIDAY_DATA;
  oscat_HOLIDAY_DATA_0_49 	: ARRAY [0..49] OF oscat_HOLIDAY_DATA;
END_TYPE

FUNCTION DAY_OF_DATE:DINT
	VAR_INPUT
		IDATE :	UDINT;
	END_VAR

	day_of_date := UDINT_TO_DINT(idate / UDINT#86400);
END_FUNCTION

FUNCTION YEAR_OF_DATE:INT
	VAR_INPUT
		IDATE :	UDINT;
	END_VAR

	YEAR_OF_DATE := UDINT_TO_INT((idate+UDINT#43200) / UDINT#31557600 + UDINT#1970);
END_FUNCTION

FUNCTION _INT_TO_UDINT:UDINT
	VAR_INPUT
		IN :	INT;
	END_VAR

	_INT_TO_UDINT := DINT_TO_UDINT(INT_TO_DINT(IN));
END_FUNCTION

FUNCTION SET_DATE:UDINT

	VAR_INPUT
		YEAR :	INT;
		MONTH :	INT;
		DAY :	INT;
	END_VAR

	VAR
		count :	INT;
	END_VAR

	IF month > 2 THEN
		count := (month - 1) * 30;
		IF month > 7 THEN
			count := count + DWORD_TO_INT(SHR(DINT_TO_DWORD(INT_TO_DINT(month) - INT_TO_DINT(3)),1));
		ELSE
			count := count + DWORD_TO_INT(SHR(DINT_TO_DWORD(INT_TO_DINT(month) - INT_TO_DINT(4)),1));
		END_IF;
		IF SHL(INT_TO_WORD(year),14) = WORD#0 THEN
			count := count + 1;
		END_IF;
	ELSE
		count := (month - 1) * 31;
	END_IF;
	SET_DATE := (_INT_TO_UDINT(count + day - 1) + DWORD_TO_UDINT(SHR(UDINT_TO_DWORD(_INT_TO_UDINT(year) * UDINT#1461 - UDINT#2878169), 2))) * UDINT#86400;
END_FUNCTION

FUNCTION_BLOCK EVENTS
	VAR_INPUT
		DATE_IN :	UDINT;
		ENA :	BOOL;
	END_VAR

	VAR_OUTPUT
		Y :	BOOL;
		NAME :	STRING;
	END_VAR

	VAR_IN_OUT
		ELIST :	oscat_HOLIDAY_DATA_0_49;
	END_VAR

	VAR
		i :	INT;
		last_active :	UDINT;
		size :	INT := 49;
		day_in :	DINT;
		cyr :	INT;
		lday :	DINT;
		check :	oscat_HOLIDAY_DATA;
		y_int :	BOOL;
		name_int :	STRING;
	END_VAR

	IF last_active <> date_in THEN
		last_active := DATE_IN;
		Y_int := FALSE;
		name_int := '';
		day_in := DAY_OF_DATE(DATE_IN);
		cyr := YEAR_OF_DATE(DATE_IN);

		(* search list for events *)
		FOR i := 0 TO size DO
			check := elist[i];
			lday := DAY_OF_DATE(SET_DATE(cyr,SINT_TO_INT(check.month), SINT_TO_INT(check.day)));
			IF day_in >= lday AND day_in <= lday + SINT_TO_DINT(check.use) - DINT#1 THEN
				y_int := TRUE;
				name_int := check.name;
				EXIT;
			END_IF;
		END_FOR;
	END_IF;

	IF ENA THEN
		Y := y_int;
		NAME := name_int;
	ELSE
		Y := FALSE;
		NAME := '';
	END_IF;

END_FUNCTION_BLOCK

PROGRAM program0
	VAR
		DATE_IN :	UDINT;
		ENA :	BOOL;

		Y :	BOOL;
		NAME :	STRING;

		ELIST :	oscat_HOLIDAY_DATA_0_49;

		func_block : EVENTS;
	END_VAR
	func_block.DATE_IN := DATE_IN;
	func_block.ENA := ENA;
	func_block.ELIST := ELIST ;

	func_block();
	Y  := func_block.Y;
	NAME  := func_block.NAME;
	ELIST  := func_block.ELIST;
END_PROGRAM

CONFIGURATION Config0
	RESOURCE Res0 ON PLC
		TASK task0(INTERVAL := T#20ms,PRIORITY := 0);
		PROGRAM instance0 WITH task0 : program0;
	END_RESOURCE
END_CONFIGURATION

(* ---- F_LAMP.ST ---- *)
FUNCTION_BLOCK T_PLC_MS_block
	VAR_OUTPUT
		T_PLC_MS :	UDINT;
	END_VAR

	VAR_EXTERNAL
		PLC_TICKS_PER_SEC :	INT;
		PLC_SYS_TICK_CNT :	DINT;
	END_VAR

	VAR
		debug :	BOOL;(*Debug-Mode ON / OFF*)
		N :	INT;(*Debug-Faktor*)
		Offset :	UDINT;(*Debug-Offset*)
		temp :	DWORD := DWORD#1;(*Debug-Offset*)
		mode :	BOOL;(*modus*)
		faktor :	UDINT;(*Systemtakt-Faktor*)
		init :	BOOL;
		v_plc_ticks_per_sec :	UDINT;
		base :	UDINT := UDINT#1000;
	END_VAR

	IF init = FALSE THEN
		v_plc_ticks_per_sec := INT_TO_UDINT(PLC_TICKS_PER_SEC);
		IF v_plc_ticks_per_sec = UDINT#1024 THEN
			faktor := UDINT#1;
			mode := FALSE;
		ELSIF v_plc_ticks_per_sec > UDINT#0 THEN
			IF v_plc_ticks_per_sec <= base THEN
				faktor := base / v_plc_ticks_per_sec;
				mode := FALSE;
			ELSE
				faktor := v_plc_ticks_per_sec / base;
				mode := TRUE;
			END_IF;
		ELSE
			faktor := UDINT#1;
		END_IF;
		init := TRUE;
	END_IF;

	IF mode THEN
		T_PLC_MS := DINT_TO_UDINT(PLC_SYS_TICK_CNT) / faktor;
	ELSE
		T_PLC_MS := DINT_TO_UDINT(PLC_SYS_TICK_CNT) * faktor;
	END_IF;

	IF debug THEN
		T_PLC_MS := (DWORD_TO_UDINT(SHL(UDINT_TO_DWORD(T_PLC_MS),N) OR SHL(temp,N)) - UDINT#1) + Offset;
	END_IF;

END_FUNCTION_BLOCK

FUNCTION_BLOCK ONTIME_Block

	VAR_INPUT
		IN :	BOOL;
		RST :	BOOL;
	END_VAR

	VAR_IN_OUT
		SECONDS :	UDINT;
		CYCLES :	UDINT;
	END_VAR

	VAR
		tx :	UDINT;
		last :	UDINT;
		edge :	BOOL;
		init :	BOOL;
		ms :	UDINT;
		T_PLC_MS :	T_PLC_MS_Block;
	END_VAR

	T_PLC_MS();
	tx:= T_PLC_MS.T_PLC_MS;

	IF NOT init THEN
		init := TRUE;
		last := tx;
		ms := UDINT#0;
	END_IF;
	IF RST THEN
		SECONDS := UDINT#0;
		CYCLES := UDINT#0;
		last := tx;
		ms := UDINT#0;
	ELSIF IN THEN
		(* add the current milliseconds *)
		ms := (tx - last) + ms;
		IF ms >= UDINT#1000 THEN
			seconds := seconds + UDINT#1;
			ms := ms - UDINT#1000;
		END_IF;
		cycles := cycles + BOOL_TO_UDINT(NOT edge);
	END_IF;
	last := tx;
	edge := in;

END_FUNCTION_BLOCK

FUNCTION_BLOCK F_LAMP_Block

	VAR_INPUT
		SWITCH :	BOOL;
		DIMM :	BYTE := BYTE#255;
		RST :	BOOL;
		T_NO_DIMM :	UINT := UINT#100;
		T_MAINTENANCE :	UINT := UINT#15000;
	END_VAR

	VAR_OUTPUT
		LAMP :	BYTE;
		STATUS :	BYTE;
	END_VAR

	VAR_IN_OUT
		ONTIME :	UDINT;
		CYCLES :	UDINT;
	END_VAR

	VAR
		runtime :	ONTIME_Block;
	END_VAR

	runtime(in := switch, SECONDS := ONTIME , CYCLES := CYCLES);
	CYCLES := runtime.CYCLES;
	ONTIME := runtime.SECONDS;

	IF RST THEN
		ONTIME := UDINT#0;
		CYCLES := UDINT#0;
	END_IF;
	IF SWITCH THEN
		IF ontime < UINT_TO_UDINT(T_NO_DIMM) * UDINT#3600 THEN
			LAMP := BYTE#255;
			STATUS := BYTE#111;
		ELSE
			LAMP := DIMM;
			STATUS := BYTE#112;
		END_IF;
	ELSE
		LAMP := BYTE#0;
		STATUS := BYTE#110;
	END_IF;

	IF ontime >= UINT_TO_UDINT(T_maintenance) * UDINT#3600 AND T_Maintenance > UINT#0 THEN
		STATUS := BYTE#120;
	END_IF;

END_FUNCTION_BLOCK

PROGRAM program0
	VAR
	    SWITCH :	BOOL;
		DIMM :	BYTE := BYTE#255;
		RST :	BOOL;
		T_NO_DIMM :	UINT := UINT#100;
		T_MAINTENANCE :	UINT := UINT#15000;
		ONTIME :	UDINT;
		CYCLES :	UDINT;
		LAMP :	BYTE;
		STATUS :	BYTE;

		func_block : F_LAMP_Block;
  	END_VAR
	func_block.SWITCH := SWITCH;
	func_block.DIMM := DIMM;
	func_block.RST := RST;
	func_block.T_NO_DIMM := T_NO_DIMM;
	func_block.T_MAINTENANCE := T_MAINTENANCE;
	func_block.ONTIME := ONTIME;
	func_block.CYCLES := CYCLES;

	func_block();
	ONTIME := func_block.ONTIME;
	CYCLES := func_block.CYCLES;
	LAMP := func_block.LAMP;
	STATUS := func_block.STATUS;
END_PROGRAM

CONFIGURATION Config0
	VAR_GLOBAL
		PLC_TICKS_PER_SEC :	INT;
		PLC_SYS_TICK_CNT :	DINT;
	END_VAR
  	RESOURCE Res0 ON PLC
    	TASK task0(INTERVAL := T#20ms,PRIORITY := 0);
    	PROGRAM instance0 WITH task0 : program0;
  	END_RESOURCE
END_CONFIGURATION

(* ---- F_POLY.ST ---- *)
TYPE
  oscat_arr_0_7               : ARRAY [0..7]    OF REAL;
END_TYPE

FUNCTION_BLOCK F_POLY_Block
	VAR_INPUT
		X :	REAL;
		C :	oscat_arr_0_7;
	END_VAR

	VAR_OUTPUT
		F_POLY :	REAL;
	END_VAR

	F_POLY := ((((((( c[7] * x + c[6] ) * x + c[5] ) * x + c[4] ) * x + c[3] ) * x + c[2] ) * x + c[1] ) * x + c[0] ) ;

END_FUNCTION_BLOCK

PROGRAM program0
	VAR
		X :	REAL;
		C :	oscat_arr_0_7;

		F_POLY :	REAL;

		func_block : F_POLY_Block;
	END_VAR
	func_block.X := X;
	func_block.C := C;
	func_block();
	F_POLY  := func_block.F_POLY;
END_PROGRAM

CONFIGURATION Config0
	RESOURCE Res0 ON PLC
		TASK task0(INTERVAL := T#20ms,PRIORITY := 0);
		PROGRAM instance0 WITH task0 : program0;
	END_RESOURCE
END_CONFIGURATION
